(* IEC 61131-3 sources: traffic-lights/PLC_TrafficLights/Class/SafetyManager (part 4) *)

          pHelpSafety^.pThis^.NewInst(pPara, pResult);

          IsDestDomain := TRUE;
          return;
        end_if;

        pHelpSafety := pHelpSafety^.pNext;
      end_while;
    end_if;
  end_if;

END_FUNCTION

FUNCTION SafetyManager::PDOLengthCorrection
  VAR
    pHelpConfig : ^t_CfgListElem;
    pHelpPDO    : ^t_PdoListElem;
    pHelpModule : ^t_ModuleListElem;
    pHelpSearchConfig : ^t_CfgListElem;
    FoundIt : BOOL;
    GotFirst : BOOL;
  END_VAR

  // with FSoE we use connections instead of the PDOs (PDOs are only remembered to check the optional state)
  if b_GotFSoEModules then
    return;
  end_if;

  GotFirst := FALSE;

  // check if there is a PDO with a zero length
  pHelpConfig := pConfigs;
  while pHelpConfig do
    pHelpPDO := pHelpConfig^.pFirstPdoCfg;
    while pHelpPDO do
      // remember the first PDO found as our act (to start from)
      if GotFirst = FALSE then
        GotFirst := TRUE;

        pActualSendCfg := pHelpConfig;
        pActualSendPDO := pHelpPDO;
      end_if;

      // if there is a PDO with no length
      if pHelpPDO^.PdoInfo.PdoLen = 0 then
        FoundIt := FALSE;
        pHelpSearchConfig := pConfigs;
        // search for the source module, because we use the length of it
        while pHelpSearchConfig & (FoundIt = FALSE) do
          pHelpModule := pHelpSearchConfig^.pFirstModuleCfg;
          while pHelpModule & (FoundIt = FALSE) do
            if pHelpModule^.ModuleInfo.PathLen = pHelpPDO^.PdoInfo.SourcePathLen then
              if (To_StdLib.MemCmp(pHelpModule^.ModuleInfo.pPath, pHelpPDO^.PdoInfo.pSourcePath, pHelpModule^.ModuleInfo.PathLen) = 0) then
                pHelpPDO^.PdoInfo.PdoLen := pHelpModule^.ModuleInfo.PdoOutLen;
                FoundIt := TRUE;
              end_if;
            end_if;

            pHelpModule := pHelpModule^.pNext;
          end_while;

          pHelpSearchConfig := pHelpSearchConfig^.pNext;
        end_while;
      end_if;

      pHelpPDO := pHelpPDO^.pNext;
    end_while;

    pHelpConfig := pHelpConfig^.pNext;
  end_while;

END_FUNCTION

FUNCTION SafetyManager::DoublePDOEntry
  VAR_INPUT
    NewPDO 	: t_PdoCfg;
    pNewCfg 	: ^t_CfgListElem;
  END_VAR
  VAR_OUTPUT
    IsDoubleEntry 	: BOOL;
  END_VAR
  VAR
    pHelpCfg : ^t_CfgListElem;
    pHelpPdo : ^t_PdoListElem;
  END_VAR

  IsDoubleEntry := FALSE;

  // if it's our first config, there is no chance for a double PDO => check only if not first config
  if pNewCfg <> pConfigs then
    // otherwise: search all prior configs for the same PDO (source and destination path match)
    pHelpCfg := pConfigs;
    while pHelpCfg <> pNewCfg do
      pHelpPdo := pHelpCfg^.pFirstPdoCfg;
      while pHelpPdo do
        if (pHelpPdo^.PdoInfo.SourcePathLen = NewPDO.SourcePathLen) & (pHelpPdo^.PdoInfo.DestPathLen = NewPDO.DestPathLen) &
           (To_StdLib.MemCmp(pHelpPdo^.PdoInfo.pSourcePath, NewPDO.pSourcePath, NewPDO.SourcePathLen) = 0) &
           (To_StdLib.MemCmp(pHelpPdo^.PdoInfo.pDestPath, NewPDO.pDestPath, NewPDO.DestPathLen) = 0) then
          // we found the same PDO in a prior config
          IsDoubleEntry := TRUE;
          return;
        end_if;

        pHelpPdo := pHelpPdo^.pNext;
      end_while;

      pHelpCfg := pHelpCfg^.pNext;
    end_while;
  end_if;

END_FUNCTION

FUNCTION SafetyManager::StoreInterfaceRoutingList
  VAR_INPUT
    pPara 	: ^CmdStruct;
    pResult 	: ^results;
    IsFSoE 	: BOOL;
  END_VAR
  VAR
    pHelpManaging : ^t_ManagingComponent;
    EntryNo       : USINT;
    i             : UDINT;
    pHelp         : ^t_InterfaceFrameInfo;
    ActOffset     : UDINT;
    pHelpFSoE     : ^t_IFConnectionInfo;
    j             : UDINT;
    GenerateNo    : USINT;
    OldFSoENo     : DINT;
  END_VAR

  if IsFSoE then

    // if we already have different data from this management component => delete the old stuff first
    if IFFSoENo then
      OldFSoENo := IFFSoENo$DINT;

      // remove the existing stuff of this managing component
      for i$DINT := (OldFSoENo-1) to 0 by -1 do
        // check if it's from the same managing component
        if aIFFSoEInfos[i].pManaging^.pThis$DINT = pPara^.aPara[2] then
          // remove it

          // move the following blocks over this one (if it's not the last)
          if i$UDINT < IFFSoENo-1 then
            for j := i to (IFFSoENo-2) do
              aIFFSoEInfos[j] := aIFFSoEInfos[j+1];
            end_for;
          end_if;
          IFFSoENo -= 1;
        end_if;
      end_for;
    end_if;

    EntryNo := ((pPara^.aPara[0] - sizeof(t_IFInfoFSoE.IsResponse)) / sizeof(t_IFConnectionInfo))$USINT;
    if (EntryNo + IFFSoENo <= MAX_MODULES_IN_OTHER_DOMAINS) then
      ActOffset := 0;
      pHelpManaging := pFirstManagingInterfaceComponent;
      while pHelpManaging do
        // if we found the sender of this list in our list of interfaceframe components, remember the safety numbers
        if pHelpManaging^.pThis$DINT = pPara^.aPara[2] then
          if EntryNo then

            // set the help pointer to the first entry of the interface frame info array
            pHelpFSoE := pPara^.aPara[1]$^t_IFConnectionInfo + sizeof(BOOL);
            for i := 0 to (EntryNo-1) do
              pHelpManaging^.ModuleInfo[i].SafetyNbr := pHelpFSoE^.SafetyNbr;

              if pHelpFSoE^.Flags.IsMaster then
                pHelpManaging^.ModuleInfo[i].InfoBits.IsFSoEMaster := TRUE;
                pHelpManaging^.ModuleInfo[i].InfoBits.IsFSoESlave  := FALSE;
              else
                pHelpManaging^.ModuleInfo[i].InfoBits.IsFSoEMaster := FALSE;
                pHelpManaging^.ModuleInfo[i].InfoBits.IsFSoESlave  := TRUE;
              end_if;

              // we save the whole info for PDO/SDO routing
              aIFFSoEInfos[IFFSoENo].FromOtherSide := pHelpFSoE^;
              aIFFSoEInfos[IFFSoENo].FromOtherSide.FollowUps := 0; // only relevant for the transfer to this domain
              aIFFSoEInfos[IFFSoENo].pManaging := pHelpManaging;

              IFFSoENo += 1;

              if pHelpFSoE^.FollowUps then
                GenerateNo := pHelpFSoE^.FollowUps;
                for j := 1 to GenerateNo do
                  // we save the whole info for PDO/SDO routing
                  aIFFSoEInfos[IFFSoENo].FromOtherSide := pHelpFSoE^;
                  aIFFSoEInfos[IFFSoENo].FromOtherSide.FollowUps := 0; // only relevant for the transfer to this domain
                  aIFFSoEInfos[IFFSoENo].pManaging := pHelpManaging;

                  IFFSoENo += 1;
                end_for;
              end_if;

              pHelpFSoE += sizeof(t_IFConnectionInfo);
            end_for;
          end_if;

          pHelpManaging^.ModuleNo := EntryNo;

          pHelpManaging^.InfoBits.GotIFInfo := TRUE;
          return;
        end_if;

        pHelpManaging := pHelpManaging^.pNext;
      end_while;
    else
      LogError("@0473 (SafetyManager::StoreInterfaceRoutingList) Invalid size of configuration (FSoE)");
    end_if;
  else
    EntryNo := ((pPara^.aPara[0] - sizeof(t_IFInfo.IsResponse)) / sizeof(t_InterfaceFrameInfo))$USINT;

    if (EntryNo + InterfaceFrameNo <= MAX_MODULES_IN_OTHER_DOMAINS) then
      ActOffset := 0;
      pHelpManaging := pFirstManagingInterfaceComponent;
      while pHelpManaging do
        // if we found the sender of this list in our list of interfaceframe components, remember the safety numbers
        if pHelpManaging^.pThis$DINT = pPara^.aPara[2] then
          if EntryNo then
            // set the help pointer to the first entry of the interface frame info array
            pHelp := pPara^.aPara[1]$^t_InterfaceFrameInfo + sizeof(BOOL);
            for i := 0 to (EntryNo-1) do
              // we save the module info's with the domain interface module for TDO/SDO routing
              pHelpManaging^.ModuleInfo[i] := pHelp^.ModuleInfo;

              // we also save the whole info for PDO routing
              aInterfaceFrameInfos[InterfaceFrameNo] := pHelp^;

              // only for IFs where the communication partner is the source
              if aInterfaceFrameInfos[InterfaceFrameNo].IFPdoLen then
                aInterfaceFrameInfos[InterfaceFrameNo].OffsetInDomainModule := ActOffset;
                ActOffset += aInterfaceFrameInfos[InterfaceFrameNo].IFPdoLen;
              end_if;

              InterfaceFrameNo += 1;

              pHelp += sizeof(t_InterfaceFrameInfo);
            end_for;
          end_if;

          pHelpManaging^.ModuleNo := EntryNo;

          pHelpManaging^.InfoBits.GotIFInfo := TRUE;
          return;
        end_if;

        pHelpManaging := pHelpManaging^.pNext;
      end_while;
    else
      LogError("@0475 (SafetyManager::StoreInterfaceRoutingList) Invalid size of configuration");
    end_if;
  end_if;

END_FUNCTION

FUNCTION SafetyManager::AllInterfaceCfgsArrived
  VAR_OUTPUT
    AllReady 	: BOOL;
  END_VAR
  VAR
    pHelpManaging : ^t_ManagingComponent;
  END_VAR

  AllReady := TRUE;

  // check if we have the safety numbers for every interface managing module in the system
  pHelpManaging := pFirstManagingInterfaceComponent;
  while pHelpManaging do
    if pHelpManaging^.InfoBits.IsSynchron & (pHelpManaging^.InfoBits.GotIFInfo = FALSE) then
      AllReady := FALSE;
      return;
    end_if;

    pHelpManaging := pHelpManaging^.pNext;
  end_while;

END_FUNCTION

FUNCTION SafetyManager::SendInterfaceConfigs
  VAR_INPUT
    DestinationThis 	: pVirtualBase;(* := NIL *)
    IsResponse 	: BOOL;(* := FALSE *)
    IsFSoE 	: BOOL;
  END_VAR
  VAR
    pHelpCfg                  : ^t_CfgListElem;
    pHelpModule               : ^t_ModuleListElem;
    pHelpPdo                  : ^t_PdoListElem;
    pHelpConnection           : ^t_FSoEConnectionDetails;
    MyPara                    : CmdStruct;
    MyResult                  : results;
    TmpIFInfo                 : t_IFInfo;
    ModuleInfoNo              : USINT;
    i                         : UDINT;
    pActCRC                   : ^HDINT;
    TmpIFConn                 : t_IFInfoFSoESend;
    pLastReferenceConnection  : ^t_IFConnectionInfo;
  END_VAR

  // collect the safety numbers of this system
  ModuleInfoNo := 0;

  if IsFSoE then
    //reset memory => now 0 is an invalid safety number (= unused element of the array)
    _memset(dest:=#TmpIFConn, usByte:=0, cntr:=sizeof(t_IFInfoFSoESend));
    TmpIFConn.IsResponse := IsResponse;

    pLastReferenceConnection  := NIL;

    // if not all configs available, create and send the available data
    if (LocalCPUCfgNo <> LocalCPUNo) then
      // check FSoE Connections in the available configs
      pHelpCfg := pConfigs;
      while pHelpCfg do
        pHelpConnection := pHelpCfg^.pFirstFSoEConnection;
        while pHelpConnection do
          // only interface connections are relevant
          if pHelpConnection^.Flags.IsInterfaceConnection then
            if pLastReferenceConnection & (pHelpConnection^.SlaveAddress = pLastReferenceConnection^.SlaveAddress) &
               (pHelpConnection^.Flags.IsMaster = pLastReferenceConnection^.Flags.IsMaster) then
              pLastReferenceConnection^.FollowUps += 1;
            else
              // add the modules to the info message
              TmpIFConn.aConnectionInfos[ModuleInfoNo].Flags            := pHelpConnection^.Flags;
              TmpIFConn.aConnectionInfos[ModuleInfoNo].SlaveAddress     := pHelpConnection^.SlaveAddress;
              TmpIFConn.aConnectionInfos[ModuleInfoNo].SafetyNbr        := pHelpConnection^.OwnerSafetyNbr;
              TmpIFConn.aConnectionInfos[ModuleInfoNo].MasterReadSize   := pHelpConnection^.MasterReadSize;
              TmpIFConn.aConnectionInfos[ModuleInfoNo].MasterWriteSize  := pHelpConnection^.MasterWriteSize;
              TmpIFConn.aConnectionInfos[ModuleInfoNo].FollowUps        := 0;

              // some data are only available at the master
              if pHelpConnection^.Flags.IsMaster then
                // no follow ups for master connections
                pLastReferenceConnection                                := NIL;

                TmpIFConn.aConnectionInfos[ModuleInfoNo].ConnectionID   := pHelpConnection^.ConnectionID;
              else
                // update this value for the next connections with the same settings to save a lot of memory
                pLastReferenceConnection                                := #TmpIFConn.aConnectionInfos[ModuleInfoNo];

                TmpIFConn.aConnectionInfos[ModuleInfoNo].ConnectionID   := 0;
              end_if;

              if pHelpConnection^.SlavePathCompLen & pHelpConnection^.pSlavePathComp then
                TmpIFConn.aConnectionInfos[ModuleInfoNo].InterfaceCRC := (pHelpConnection^.pSlavePathComp$^HDINT + 1)^;
              else
                TmpIFConn.aConnectionInfos[ModuleInfoNo].InterfaceCRC := 0;
              end_if;

              ModuleInfoNo += 1;
            end_if;
          end_if;

          pHelpConnection := pHelpConnection^.pNext;
        end_while;

        pHelpCfg := pHelpCfg^.pNext;
      end_while;
    else
      // check FSoE Connections in the sorted list
      pHelpConnection := pSortedConnections;
      while pHelpConnection do
        // only interface connections are relevant
        if pHelpConnection^.Flags.IsInterfaceConnection then
          if pLastReferenceConnection & (pHelpConnection^.SlaveAddress = pLastReferenceConnection^.SlaveAddress) &
             (pHelpConnection^.Flags.IsMaster = pLastReferenceConnection^.Flags.IsMaster) then
            pLastReferenceConnection^.FollowUps += 1;
          else
            // add the modules to the info message
            TmpIFConn.aConnectionInfos[ModuleInfoNo].Flags            := pHelpConnection^.Flags;
            TmpIFConn.aConnectionInfos[ModuleInfoNo].SlaveAddress     := pHelpConnection^.SlaveAddress;
            TmpIFConn.aConnectionInfos[ModuleInfoNo].SafetyNbr        := pHelpConnection^.OwnerSafetyNbr;
            TmpIFConn.aConnectionInfos[ModuleInfoNo].MasterReadSize   := pHelpConnection^.MasterReadSize;
            TmpIFConn.aConnectionInfos[ModuleInfoNo].MasterWriteSize  := pHelpConnection^.MasterWriteSize;
            TmpIFConn.aConnectionInfos[ModuleInfoNo].FollowUps        := 0;

            // some data are only available at the master
            if pHelpConnection^.Flags.IsMaster then
              // no follow ups for master connections
              pLastReferenceConnection                                := NIL;

              TmpIFConn.aConnectionInfos[ModuleInfoNo].ConnectionID   := pHelpConnection^.ConnectionID;
            else
              // update this value for the next connections with the same settings to save a lot of memory
              pLastReferenceConnection                                := #TmpIFConn.aConnectionInfos[ModuleInfoNo];

              TmpIFConn.aConnectionInfos[ModuleInfoNo].ConnectionID   := 0;
            end_if;

            if pHelpConnection^.SlavePathCompLen & pHelpConnection^.pSlavePathComp then
              TmpIFConn.aConnectionInfos[ModuleInfoNo].InterfaceCRC := (pHelpConnection^.pSlavePathComp$^HDINT + 1)^;
            else
              TmpIFConn.aConnectionInfos[ModuleInfoNo].InterfaceCRC := 0;
            end_if;

            ModuleInfoNo += 1;
          end_if;
        end_if;

        pHelpConnection := pHelpConnection^.pNextSorted;
      end_while;
    end_if;

    CheckLocalSlaveAddresses();

    if b_AllLocalSlaveAddressesValid then
      MyPara.uiCmd := CMD_SM_IF_MODULE_INFO_FSOE_OK;
    else
      MyPara.uiCmd := CMD_SM_IF_MODULE_INFO_FSOE;
    end_if;

    MyPara.aPara[0] := ModuleInfoNo * sizeof(t_IFConnectionInfo) + sizeof(t_IFInfoFSoE.IsResponse);
    MyPara.aPara[1] := (#TmpIFConn)$DINT;
  else
    // browse through the configs
    TmpIFInfo.IsResponse := IsResponse;

    pHelpCfg := pConfigs;
    while pHelpCfg do
      pHelpPdo := pHelpCfg^.pFirstPdoCfg;
      while pHelpPdo do
        // if it's a interface broadcast
        if pHelpPdo^.PdoInfo.Info.IFBroadCast then
          // search for the source module
          pHelpModule := pHelpCfg^.pFirstModuleCfg;
          while pHelpModule do
            // if it's an interface source and the interface CRC matches the one of our PDO => Bingo! But to be sure we check also the path length and the path itself
            if pHelpModule^.ModuleInfo.Info.IsInterfaceSource & (pHelpModule^.ModuleInfo.InterfaceCRC = pHelpPdo^.PdoInfo.InterfaceCRC) &
              (pHelpModule^.ModuleInfo.PathLen = pHelpPdo^.PdoInfo.SourcePathLen) &
              (To_StdLib.MemCmp(pHelpModule^.ModuleInfo.pPath, pHelpPdo^.PdoInfo.pSourcePath, pHelpPdo^.PdoInfo.SourcePathLen) = 0) then

              TmpIFInfo.aModuleInfos[ModuleInfoNo].InterfaceCRC          := pHelpModule^.ModuleInfo.InterfaceCRC;
              TmpIFInfo.aModuleInfos[ModuleInfoNo].IFPdoLen              := pHelpPdo^.PdoInfo.PdoLen;
              TmpIFInfo.aModuleInfos[ModuleInfoNo].OffsetInDomainModule  := 0; // the correct offset is calculated in the receiver
              TmpIFInfo.aModuleInfos[ModuleInfoNo].ModuleInfo.SafetyNbr  := pHelpModule^.ModuleInfo.SafetyNbr;

              ModuleInfoNo += 1;
            end_if;

            pHelpModule := pHelpModule^.pNext;
          end_while;
        end_if;

        pHelpPdo := pHelpPdo^.pNext;
      end_while;

      // check the modules of the actual config if there are interface frame destinations (needed for unidirectional communication, otherwise the SDO routing would fail)
      pHelpModule := pHelpCfg^.pFirstModuleCfg;
      while pHelpModule do
        // if it's a interface destination
        if pHelpModule^.ModuleInfo.Info.IsInterfaceDest then
          pActCRC := pHelpModule^.ModuleInfo.pDestCRCs;
          for i := 0 to (pHelpModule^.ModuleInfo.DestCRCNo-1) do
            TmpIFInfo.aModuleInfos[ModuleInfoNo].InterfaceCRC          := pActCRC^;
            TmpIFInfo.aModuleInfos[ModuleInfoNo].IFPdoLen              := 0; // we don't know the length here, we're only the receiver
            TmpIFInfo.aModuleInfos[ModuleInfoNo].OffsetInDomainModule  := 0; // the correct offset is calculated in the receiver
            TmpIFInfo.aModuleInfos[ModuleInfoNo].ModuleInfo.SafetyNbr  := pHelpModule^.ModuleInfo.SafetyNbr;
            TmpIFInfo.aModuleInfos[ModuleInfoNo].ModuleInfo.InfoBits$UDINT := 0;

            pActCRC += sizeof(HDINT);
            ModuleInfoNo += 1;
          end_for;
        end_if;

        pHelpModule := pHelpModule^.pNext;
      end_while;

      pHelpCfg := pHelpCfg^.pNext;
    end_while;

    MyPara.uiCmd := CMD_SM_IF_MODULE_INFO;
    MyPara.aPara[0] := ModuleInfoNo * sizeof(t_InterfaceFrameInfo) + sizeof(TmpIFInfo.IsResponse);
    MyPara.aPara[1] := (#TmpIFInfo)$DINT;
  end_if;

  // if we have only 1 destination => sent it to this destination
  if DestinationThis then
    DestinationThis^.NewInst(#MyPara, #MyResult);
  else
    // otherwise send our safety numbers to every interface managing module in the system
    TellAllInterfaceManagingModules(#MyPara, #MyResult);
  end_if;

END_FUNCTION

FUNCTION SafetyManager::GetIFInfoByCRC
  VAR_INPUT
    InterfaceCRC 	: HDINT;
    pMemOffset 	: ^UDINT;
    pLength 	: ^USINT;
  END_VAR
  VAR_OUTPUT
    SafetyNbr 	: HDINT;
  END_VAR
  VAR
    i : UDINT;
  END_VAR

  SafetyNbr := 0;

  if InterfaceFrameNo then
    for i := 0 to (InterfaceFrameNo-1) do
      // if we found the interface CRC and it's a interface frame we receive (the sender adds the length)
      if (aInterfaceFrameInfos[i].InterfaceCRC = InterfaceCRC) & aInterfaceFrameInfos[i].IFPdoLen then
        SafetyNbr := aInterfaceFrameInfos[i].ModuleInfo.SafetyNbr;
        // check if pointers are valid
        if pMemOffset & pLength then
          pMemOffset^ := aInterfaceFrameInfos[i].OffsetInDomainModule;
          pLength^    := aInterfaceFrameInfos[i].IFPdoLen;
        end_if;
        return;
      end_if;
    end_for;

    if SafetyNbr = 0 then
      LogError("@0476 (SafetyManager::GetIFInfoByCRC) Safetynumber of Interface-Frame source couldn't be found in the list");
    end_if;
  end_if;

END_FUNCTION

FUNCTION SafetyManager::SetTimeout

  ud_InitTimeOut := ops.tAbsolute;

END_FUNCTION

FUNCTION SafetyManager::CheckTimeout

  // if the step took too long
  if (OPS.tAbsolute - ud_InitTimeOut) > T_INIT_TIMEOUT then
    // show the possible error in the log/trace and restart the time for timeout
    case InitSSW of
//**********************************************************************************************************************************************************
      _FirstWait4SynchronSubdomains:
        LogError("@0477 (SafetyManager::CheckTimeout) Timeout in Initialisation while waiting first time for subdomains to get synchron!");
//**********************************************************************************************************************************************************
      _Wait4FSoEConnectionsLocal:
        LogError("@0478 (SafetyManager::CheckTimeout) Timeout in Initialisation while waiting for the local FSoE connections to get initialized!");
//**********************************************************************************************************************************************************
      _Wait4SynchronSubdomains:
        LogError("@0479 (SafetyManager::CheckTimeout) Timeout in Initialisation while waiting for subdomains to get synchron!");
//**********************************************************************************************************************************************************
//      _Wait4ConfigFlush:
//        LogError("@ZZZZ Timeout in Initialisation while waiting for the slave domains to send their safety numbers of safety cpus and if they can handle the new time sync method!");
//**********************************************************************************************************************************************************
      _Wait4CPUConfigs:
        LogError("@047A (SafetyManager::CheckTimeout) Timeout in Initialisation while waiting for all available cpu configurations!");
//**********************************************************************************************************************************************************
      _Wait4InterfaceConfigs:
        LogError("@047B (SafetyManager::CheckTimeout) Timeout in Initialisation while waiting for module info needed for interface frame communication!");
//**********************************************************************************************************************************************************
      _Wait4FSoEConnectionsExternal:
        LogError("@047C (SafetyManager::CheckTimeout) Timeout in Initialisation while waiting for the external FSoE connections to get initialized!");
//**********************************************************************************************************************************************************
      _Wait4UnsafeConfigAck:
        LogError("@047D (SafetyManager::CheckTimeout) Timeout in Initialisation while waiting for an unsafe variable configuration acknowledgment!");
//**********************************************************************************************************************************************************
      _Wait4PDOAcks:
        LogError("@047F (SafetyManager::CheckTimeout) Timeout in Initialisation while waiting for a pdo configuration acknowledgment!");
//**********************************************************************************************************************************************************
    end_case;

    // this error gets quitted if initialisation finishes
    ClassState := -11;

    ud_InitTimeOut := ops.tAbsolute;
  end_if;

END_FUNCTION

FUNCTION SafetyManager::AllNonOptionalIFDomainsSynchron
  VAR_OUTPUT
    EverythingSynchron 	: BOOL;
  END_VAR
  VAR
    pHelpManaging : ^t_ManagingComponent;
    pHelpConfig : ^t_CfgListElem;
    pHelpPdo : ^t_PdoListElem;
    TempCfg : t_PdoCfg;
    MyPara 	  : CmdStruct;
    MyResult	: results;
  END_VAR

  EverythingSynchron := TRUE;

  MyPara.uiCmd := CMD_SM_SYNC_CHECK;

  // check for all interface frame PDOs in the configurations if the corresponding domain managing module is synchron
  pHelpConfig := pConfigs;
  while pHelpConfig do
    pHelpPdo := pHelpConfig^.pFirstPdoCfg;
    while pHelpPdo do
      TempCfg := pHelpPdo^.PdoInfo;
      // if it's an interface  PDO, no double entry and not optional => it has to be synchron!
      if (TempCfg.Info.IsInterfacePDO = TRUE) & (TempCfg.Info.DoublePDOEntry = FALSE) & (TempCfg.Info.IsOptional = FALSE) then
        pHelpManaging := pFirstManagingInterfaceComponent;
        while pHelpManaging do
          // we found the corresponding domain managing module
          if (pHelpManaging^.InfoBits.IsOptional = FALSE) &
            ((To_StdLib.MemCmp(pHelpManaging^.pModulePath, TempCfg.pSourcePath, TempCfg.SourcePathLen) = 0) |
             (To_StdLib.MemCmp(pHelpManaging^.pModulePath, TempCfg.pDestPath, TempCfg.DestPathLen) = 0)) then

            // if any of those is not synchron, stop searching
            if pHelpManaging^.pThis^.NewInst(#MyPara, #MyResult) = ERROR then
              EverythingSynchron := FALSE;
              return;
            end_if;

            exit;
          end_if;

          pHelpManaging := pHelpManaging^.pNext;
        end_while;
      end_if;

      pHelpPdo := pHelpPdo^.pNext;
    end_while;

    pHelpConfig := pHelpConfig^.pNext;
  end_while;

END_FUNCTION

FUNCTION VIRTUAL SafetyManager::GetThisViaServerName
  VAR_INPUT
    pObjectDotServer 	: ^CHAR;
  END_VAR
  VAR_OUTPUT
    ThisPtr 	: pVoid;
  END_VAR
  VAR
    ChannelMode : CHMODE;
  END_VAR

  ThisPtr := NIL;

  if pObjectDotServer = NIL then
    return;
  end_if;

  // get thispointer to server via name
  ChannelMode := _LookUpEmbed_C(pObjectDotServer, #ThisPtr, NIL);

  // check if it's a server
  case ChannelMode of
    _CH_CMD,
    _CH_SVR:

  else
    ThisPtr := NIL;
    LogError("@0480 (SafetyManager::GetThisViaServerName) Couldn't get thispointer of server:");
    LogError(e_msg:=pObjectDotServer);
  end_case;

END_FUNCTION

FUNCTION SafetyManager::GetNewMovDO
  VAR_OUTPUT
    Index 	: INT;
  END_VAR
//  VAR
//  	sd_retval : DINT;
//  END_VAR

  Index := -1;

  if CopyCmdsUsed < MAX_PDO_COPY_CMDS then
    // check if there is one available but not used
    if CopyCmdsUsed < CopyCmdsAvailable then
      Index := CopyCmdsUsed;
      CopyCmdsUsed += 1;
    else
      // we have to create a new one

(*
// connection to varan manager required
      // add data object to copy our data
      sd_retval := pVaranManager^.AddMovDO(ud_dol_type:=VARAN_DOL_ISO
                                         , p_ud_handle:=(#aCopyCmds[CopyCmdsAvailable].pHandle)$^UDINT
                                         , p_ud_MovSettings:=( #aCopyCmds[CopyCmdsAvailable].pSettings)$^UDINT
                                         , ud_type := VM_PRIORITY_2
                                         );

      //look for an error
      if ( sd_retval <> 0 ) then
        ClassState := -9;
        LogError("@ZZZZ (SafetyManager::GetNewMovDO) Failed to add a new copy command to the VaranManager!");
        return;
      end_if;
*)
      aCopyCmds[CopyCmdsAvailable].b_Ready4Action := FALSE;

      Index := CopyCmdsAvailable;

      CopyCmdsAvailable += 1;
      CopyCmdsUsed += 1;
    end_if;
  else
    LogError("@0481 (SafetyManager::GetNewMovDO) Maximum of possible PDO copy commands reached!");
  end_if;

END_FUNCTION

FUNCTION SafetyManager::CheckCPUConfigs
  VAR_OUTPUT
    ConfigsOK 	: BOOL;
  END_VAR
  VAR
    pHelpManaging   : ^t_ManagingComponent;
    pSourceManaging : ^t_ManagingComponent;
    pHelpConfig     : ^t_CfgListElem;
    pHelpPdo        : ^t_PdoListElem;
    pLastPdo        : ^t_PdoListElem;
    IsSource        : DINT;
    PDOCount : UDINT;
  END_VAR

  // before we go into the usual check routine, we have to ensure that we have enough virtual PDOs for writing interface frames (config holds a broadcast and we have to look for possible target modules)
  CreateVirtualPDOs();

  // initialize with true (normal case is that everything is ok => now we check for errors)
  ConfigsOK := TRUE;

  PDOCount := 0;

  // check if all non-optional modules are available and all corresponding domain managing module are synchron (if necessary)
  pHelpConfig := pConfigs;
  while pHelpConfig do
    pLastPdo := NIL;
    pHelpPdo := pHelpConfig^.pFirstPdoCfg;
    while pHelpPdo do
      // if it's an interface frame and no broadcast frame
      if pHelpPdo^.PdoInfo.Info.IsInterfacePDO then
        if (pHelpPdo^.PdoInfo.Info.IFBroadCast = FALSE) then

          // check if we have already added the domain interface to the IF List
          IsSource := -1; // -1 = not found, 0 = destination, 1 = source
          pSourceManaging := NIL;
          pHelpManaging := pFirstManagingInterfaceComponent;
          while pHelpManaging do
            // if source or destination of the PDO matches our managing module path => it's an interface frame to/from this domain
            if (To_StdLib.MemCmp(pHelpManaging^.pModulePath, pHelpPdo^.PdoInfo.pSourcePath, pHelpPdo^.PdoInfo.SourcePathLen) = 0) then
              pSourceManaging := pHelpManaging;
              IsSource := 1;
              exit;
            elsif (To_StdLib.MemCmp(pHelpManaging^.pModulePath, pHelpPdo^.PdoInfo.pDestPath, pHelpPdo^.PdoInfo.DestPathLen) = 0) then
              IsSource := 0;
              exit;
            end_if;

            pHelpManaging := pHelpManaging^.pNext;
          end_while;

          // if we got a source managing module and it isn't synchron
          if pSourceManaging then
            // if this pdo is not optional => the source module also isn't
            if pHelpPdo^.PdoInfo.Info.IsOptional = FALSE then
              pSourceManaging^.InfoBits.IsOptional := FALSE;
            end_if;

            if (pSourceManaging^.InfoBits.IsSynchron = FALSE) then
              if pHelpPdo^.PdoInfo.Info.IsOptional then
                // ignore it
  //              LogError("Info: Optional interface frame can't be received, because source domain is not connected or not synchron");

                // remove the PDO from the list (if not the receiver module would wait endless for the PDO and we can't send the set bus ready to quit errors of local PDOs)
                if pLastPdo then
                  // if we had already a PDO before in this configuration we have to skip the removed PDO with the next pointer
                  pLastPdo^.pNext := pHelpPdo^.pNext;

                  To_StdLib.Free(pHelpPdo^.PdoInfo.pSourcePath);
                  To_StdLib.Free(pHelpPdo^.PdoInfo.pDestPath);
                  To_StdLib.Free(pHelpPdo);

                  pHelpPdo := pLastPdo;
                else
                  // if it was the first PDO, we have to correct the first pointer
                  pHelpConfig^.pFirstPdoCfg := pHelpPdo^.pNext;

                  To_StdLib.Free(pHelpPdo^.PdoInfo.pSourcePath);
                  To_StdLib.Free(pHelpPdo^.PdoInfo.pDestPath);
                  To_StdLib.Free(pHelpPdo);

                  pHelpPdo := pHelpConfig^.pFirstPdoCfg;
                end_if;

                if pHelpPdo = NIL then
                  exit;
                end_if;
              else
                // non-optional interface frame domain missing => error
                LogError("@0482 (SafetyManager::CheckCPUConfigs) ERROR! Non-Optional interface frame can't be received, because domain is not connected");
                ConfigsOK := FALSE;
                ClassState := -10;
              end_if;
            end_if;
          end_if;
        end_if;
      end_if;

      PDOCount += 1;

      pLastPdo := pHelpPdo;
      pHelpPdo := pHelpPdo^.pNext;
    end_while;

    pHelpConfig := pHelpConfig^.pNext;
  end_while;

  // if now PDOs found => reset the act ID to show that there are none
  if PDOCount = 0 then
    ActPDO_ID := 0;
  end_if;

END_FUNCTION

FUNCTION SafetyManager::RemoveLocalCPUCfg
  VAR_INPUT
    SafetyNumber 	: HDINT;
  END_VAR
  VAR
    pHelpCfg    : ^t_LocalCfgListElem;
    i : UDINT;
  END_VAR

  if LocalCPUCfgNo then
    pHelpCfg := pFirstLocalCPUCfg;
    for i := 0 to (LocalCPUCfgNo-1) do
      if pHelpCfg^.SafetyNbr = SafetyNumber then
        // found it => deactivate it
        pHelpCfg^.ConfigSize := 0;
        pHelpCfg^.ConfigSent2Master := FALSE;
        exit;
      end_if;

      pHelpCfg := pHelpCfg^.pNext;
    end_for;
  end_if;

END_FUNCTION

FUNCTION SafetyManager::ClearRoutingInformations
  VAR_OUTPUT
    finished 	: BOOL;
  END_VAR
  VAR
    MyPara        : CmdStruct;
    MyResult      : results;
    pHelpManaging : ^t_ManagingComponent;
    i             : UDINT;
    pHelpCfg      : ^t_LocalCfgListElem;
    pPDOElement   : ^t_PDOElement;
    pInputPDO     : ^t_InputPDOs;
    retcode       : DINT;
    pActConnection: ^t_UdpConnection;
    pUdpNo        : ^UDINT;
    paUdpCons     : ^t_aUdpConnections;
  END_VAR

  finished := FALSE;

  if sUdpVars.ProducerConnectionNo then
    pUdpNo    := #sUdpVars.ProducerConnectionNo;
    paUdpCons := sUdpVars.paConnectionsToProducers;
  elsif sUdpVars.ConsumerConnectionNo then
    pUdpNo    := #sUdpVars.ConsumerConnectionNo;
    paUdpCons := sUdpVars.paConnectionsToConsumers;
  else
    // no UDP connections => proceed to last step
    sUdpVars.ClearRoutingInfoSSW := t_ClearRoutingInfoSSW::_FinishEverythingElse;
  end_if;

  case sUdpVars.ClearRoutingInfoSSW of
//**********************************************************************************************************************************************************
    t_ClearRoutingInfoSSW::_PrepareUdpDisconnect:
      // reset all send markers, because we will need them in the next step
      pActConnection := #paUdpCons^[0];
      for i := 0 to (pUdpNo^-1) do
        pActConnection^.WaitForResponse      := FALSE;
        pActConnection^.bSequenceCntReceived := FALSE; //reset flag to allow sequence counter for new udp communication
        pActConnection^.ActReceiveData.usHeaderVersion := 0;
        pActConnection^.ActSendData.usHeaderVersion    := 0;
        pActConnection^.RequestRetries                 := 0;

        pActConnection += sizeof(t_UdpConnection);
      end_for;

      sUdpVars.ClearRoutingInfoSSW := t_ClearRoutingInfoSSW::_SendDisconnect;

//**********************************************************************************************************************************************************
    t_ClearRoutingInfoSSW::_SendDisconnect:

      // if it's the source of the reinit => don't send him the info, just remove from the list
      if (paUdpCons^[pUdpNo^-1].IP = 0) | (paUdpCons^[pUdpNo^-1].IP = sUdpVars.ReInitSenderIP) then
        pUdpNo^ -= 1;
      else
        // disconnect all UDP connections (1 by 1 or we might get a problem with the net load)
        sUdpVars.pTempSendBufferCy^.Header.Command       := t_UdpCommand::UdpCmd_ReInitialize;
        sUdpVars.pTempSendBufferCy^.Header.State         := t_UdpPacketHeaderV2.State.IsFromConsumer OR t_UdpPacketHeaderV2.State.IsFromProducer; // invalid state for normal data

        paUdpCons^[pUdpNo^-1].InfoBits.Disconnecting  := TRUE;
        paUdpCons^[pUdpNo^-1].WaitForResponse         := TRUE;
        paUdpCons^[pUdpNo^-1].TLastRequest            := ops.tAbsolute;

        // only send command and state
        retcode := SendUDPData(sUdpVars.pTempSendBufferCy, sizeof(t_UdpPacketHeaderV2.Command) + sizeof(t_UdpPacketHeaderV2.State), paUdpCons^[pUdpNo^-1].IP);

        if retcode < 0 then
          sUdpVars.LastSendError := retcode;
          sUdpVars.SendErrorCnt += 1;
        end_if;

        sUdpVars.ClearRoutingInfoSSW := t_ClearRoutingInfoSSW::_Wait4DisconnectConfirm;
      end_if;

//**********************************************************************************************************************************************************
    t_ClearRoutingInfoSSW::_Wait4DisconnectConfirm:

      // check for the confirmation
      if paUdpCons^[pUdpNo^-1].InfoBits.Disconnecting = FALSE then

        // reset the IP address of all others with the same IP to not resend if there are multiple connections to this IP
        if sUdpVars.ConsumerConnectionNo then
          pActConnection := #sUdpVars.paConnectionsToConsumers^[0];
          for i := 0 to (sUdpVars.ConsumerConnectionNo-1) do
            // check if it's the same IP
            if (pActConnection^.IP = paUdpCons^[pUdpNo^-1].IP) then
              // reset the IP
              pActConnection^.IP := 0;
            end_if;

            pActConnection += sizeof(t_UdpConnection);
          end_for;
        end_if;

        if sUdpVars.ProducerConnectionNo then
          pActConnection := #sUdpVars.paConnectionsToProducers^[0];
          for i := 0 to (sUdpVars.ProducerConnectionNo-1) do
            // check if it's the same IP
            if (pActConnection^.IP = paUdpCons^[pUdpNo^-1].IP) then
              // reset the IP
              pActConnection^.IP := 0;
            end_if;

            pActConnection += sizeof(t_UdpConnection);
          end_for;
        end_if;

        // this one is out fine => proceed with the next
        pUdpNo^ -= 1;
        sUdpVars.ClearRoutingInfoSSW := t_ClearRoutingInfoSSW::_SendDisconnect;

      // look if we actual wait for a response to send retries and check if we didn't receive data in time
      elsif (paUdpCons^[pUdpNo^-1].WaitForResponse = TRUE) & ((ops.tAbsolute - paUdpCons^[pUdpNo^-1].TLastRequest) > (sUdpVars.CalculatedRequestTimeout * 2)) then

        if paUdpCons^[pUdpNo^-1].RequestRetries >= (UDP_MAX_RETRIES * 2) then

          // we had enough retries, just forget about this one and proceed with the next
          pUdpNo^ -= 1;
          sUdpVars.ClearRoutingInfoSSW := t_ClearRoutingInfoSSW::_SendDisconnect;
        else

          //send retry to actual cpu
          paUdpCons^[pUdpNo^-1].RequestRetries += 1;
          sUdpVars.ClearRoutingInfoSSW := t_ClearRoutingInfoSSW::_SendDisconnect;
        end_if;

      end_if;

      // producer finished but still some consumer connections to go
      if (pUdpNo^ = 0) then
        if sUdpVars.ConsumerConnectionNo then
          // go back to the initialisation and do it for the consumer connections now
          sUdpVars.ClearRoutingInfoSSW := t_ClearRoutingInfoSSW::_PrepareUdpDisconnect;
        else
          // all connections disconnected => finish the rest
          sUdpVars.ClearRoutingInfoSSW := t_ClearRoutingInfoSSW::_FinishEverythingElse;
        end_if;
      end_if;

//**********************************************************************************************************************************************************
    t_ClearRoutingInfoSSW::_FinishEverythingElse:

      // we're flushin our stuff here

      // forget who sent us the reinitialize
      sUdpVars.ReInitSenderIP := 0;

      // set ID to zero for the next mapping assignment
      ActPDO_ID := 0;

      // reset interface frameno
      InterfaceFrameNo := IFFSoENo := 0;

      // reset local interface frameno
      LocalIFNo := 0;

      // clear configurations of safety-cpus
      FreeCfgLists();

      // clear number of copy DOs used
      CopyCmdsUsed := 0;

      // reset flexible constellation informations
      _memset(dest:=#sFlexCon, usByte:=0, cntr:=sizeof(t_FlexCon));

      // reset memory usage for isochronous transfer (the values are set when distributing the PDOs)
      MyPara.aPara[0] := 0;
      pHelpManaging := pFirstManagingInterfaceComponent;
      while pHelpManaging do
        pHelpManaging^.PDOReadMemUsed := 0;
        pHelpManaging^.PDOWriteMemUsed := 0;

        MyPara.uiCmd := CMD_SM_PDO_MEM_USAGE_WR;
        pHelpManaging^.pThis^.NewInst(#MyPara, #MyResult);

        MyPara.uiCmd := CMD_SM_PDO_MEM_USAGE_RD;
        pHelpManaging^.pThis^.NewInst(#MyPara, #MyResult);

        pHelpManaging^.InfoBits.HasBeenFlushed      := FALSE;
        pHelpManaging^.InfoBits.NewTimeSyncPossible := FALSE;
        pHelpManaging^.InfoBits.SubDomainsSynchron  := FALSE;
        pHelpManaging^.InfoBits.GotIFInfo           := FALSE;
        pHelpManaging^.InfoBits.LocalConfigReady    := FALSE;
        pHelpManaging^.InfoBits.IsOptional          := TRUE;  // initialize with true, later in the init process (CheckCPUConfigs) it's checked and corrected if necessary
        // synchron bit is already true at this time (or the timeout has expired)

        pHelpManaging^.DomainNr := 16#FF;

        pHelpManaging^.SubDomainsUsed := 0;
        _memset(dest:=#pHelpManaging^.SubDomainNr, usByte:=16#FF, cntr:=sizeof(pHelpManaging^.SubDomainNr));

        pHelpManaging^.ModuleNo := 0;
        _memset(dest:=#pHelpManaging^.ModuleInfo, usByte:=16#00, cntr:=sizeof(pHelpManaging^.ModuleInfo));

        // delete flexcon information
        _memset(dest:=#pHelpManaging^.FlexCon, usByte:=0, cntr:=sizeof(t_ManagingFlexCon));

        pHelpManaging := pHelpManaging^.pNext;
      end_while;

      // all local cpu configs have to be sent again on reconnect
      if LocalCPUCfgNo then
        pHelpCfg := pFirstLocalCPUCfg;
        for i := 0 to (LocalCPUCfgNo-1) do
          pHelpCfg^.ConfigSent2Master := FALSE;

          pHelpCfg := pHelpCfg^.pNext;
        end_for;
      end_if;

      if PDOElementNo then

        // at first we have to check if there are any safety modules out there with a pointer to the PDO List (if they use a VMC/VBC as source)
        pPDOElement := #aPDOElements[0];
        for i := 0 to (PDOElementNo-1) do
          if (pPDOElement^.ThisDomainsRole = SourceDest_IsDest) & (pPDOElement^.SourceInfo.pPDOMem) & (pPDOElement^.pSafety) then
            // unregister this PDO
            MyPara.uiCmd := CMD_SM_REMOVE_INPUT_PDO;
            MyPara.aPara[0] := pPDOElement^.SourceInfo.pPDOMem$DINT;
            MyPara.aPara[1] := pPDOElement^.SourceInfo.pPDOMemDPRAM$DINT;
            pPDOElement^.pSafety^.pThis^.NewInst(#MyPara, #MyResult);
          end_if;

          // free the memory of the path infos and reset the rest of pdo element info
          if pPDOElement^.SourceInfo.pPath then
            To_StdLib.Free(pPDOElement^.SourceInfo.pPath);
          end_if;
          if pPDOElement^.DestInfo.pPath then
            To_StdLib.Free(pPDOElement^.DestInfo.pPath);
          end_if;

          pPDOElement += sizeof(t_PDOElement);
        end_for;

        _memset(dest:=#aPDOElements, usByte:=0, cntr:=PDOElementNo * sizeof(t_PDOElement));
        PDOElementNo := 0;
      end_if;

      if FSoECopyCmdNo then
        _memset(dest:=#aFSoECopyCmds, usByte:=0, cntr:=FSoECopyCmdNo * sizeof(t_FSoECopyCmd));
        FSoECopyCmdNo := 0;
      end_if;

      if FSoEInputPDONo then
        pInputPDO := #aFSoEInputPDOs[0];
        for i := 0 to (FSoEInputPDONo-1) do
          // unregister this PDO
          MyPara.uiCmd := CMD_SM_REMOVE_INPUT_PDO;
          MyPara.aPara[0] := pInputPDO^.pMem;
          MyPara.aPara[1] := 0;
          pInputPDO^.pSafety^.pThis^.NewInst(#MyPara, #MyResult);

          pInputPDO += sizeof(t_InputPDOs);
        end_for;

        FSoEInputPDONo := 0;
      end_if;

      // reset other udp settings that are not directly connected to the udp connections
      sUdpVars.UdpInit.ProvidesIF            := 0; // no need to install callback twice and FSoE is still available if it was before
      sUdpVars.LowestTransmissionTime_ms  := UDP_DEFAULT_TRANSMISSION_TIME;
      sUdpVars.ConnectionsInitialized     := FALSE;

      // set scheduler to default until a connection is established
      SetUdpSchedulerGrid();

      if sUdpVars.SendCopyCmdNo then
        _memset(dest:=#sUdpVars.aSendCopyCmds, usByte:=0, cntr:=sUdpVars.SendCopyCmdNo * sizeof(t_FSoECopyCmd));
        sUdpVars.SendCopyCmdNo := 0;
      end_if;

      if sUdpVars.ReceiveCopyCmdNo then
        _memset(dest:=#sUdpVars.aReceiveCopyCmds, usByte:=0, cntr:=sUdpVars.ReceiveCopyCmdNo * sizeof(t_FSoECopyCmd));
        sUdpVars.ReceiveCopyCmdNo := 0;
      end_if;

      // reset step
      sUdpVars.ClearRoutingInfoSSW := t_ClearRoutingInfoSSW::_PrepareUdpDisconnect;

      finished := TRUE;

  end_case;

END_FUNCTION

FUNCTION SafetyManager::CheckPDORecycle
  VAR_INPUT
    SourceDest 	: t_SourceDest;
    pNewPDO 	: ^t_PDOElement;
  END_VAR
  VAR_OUTPUT
    pRecyclePDO 	: ^t_PDOElement;
  END_VAR
  VAR
    i : UDINT;
    pHelpInfo : ^t_PDOModuleInfo;
    pSearchInfo : ^t_PDOModuleInfo;
    ppHelpManaging : ^t_pManagingComponent;
    pSearchManaging : ^t_ManagingComponent;
  END_VAR

  // initialize with invalid
  pRecyclePDO := NIL;

  // if we have no pdoelements yet, quit
  if PDOElementNo = 0 then
    return;
  end_if;

  // we search for a PDO with the same source (then it contains the same data)
  pHelpInfo := #aPDOElements[0].SourceInfo;
  pSearchInfo := #pNewPDO^.SourceInfo;

  case SourceDest of
    SourceDest_IsSource:
      ppHelpManaging := #aPDOElements[0].pManagingSource;
      pSearchManaging := pNewPDO^.pManagingSource;
    SourceDest_IsDest:
      ppHelpManaging := #aPDOElements[0].pManagingDest;
      pSearchManaging := pNewPDO^.pManagingDest;
  else
    return;
  end_case;

  // check if we already have the path info of this source/destination
  for i := 0 to (PDOElementNo-1) do
    // if managing node, pathlength and path matches
    if (ppHelpManaging^ = pSearchManaging) & (pHelpInfo^.PathLen = pSearchInfo^.PathLen) & (To_StdLib.MemCmp(pHelpInfo^.pPath, pSearchInfo^.pPath, pHelpInfo^.PathLen) = 0) then
      // we found our PDO to recycle (PDO is already tranferred over this managing node
      pRecyclePDO := #aPDOElements[i];
      return;
    end_if;

    pHelpInfo       += sizeof(t_PDOElement);
    ppHelpManaging  += sizeof(t_PDOElement);
  end_for;

END_FUNCTION

FUNCTION SafetyManager::AddManagingInfo
  VAR_INPUT
    pPara 	: ^CmdStruct;
  END_VAR
  VAR
    pHelpManaging : ^t_ManagingComponent;
  END_VAR

(*
  Parameter description:
  0..pointer to write PDOs in VARAN manager DPRAM
  1..pointer to read PDOs in VARAN manager DPRAM
  2..thispointer of calling class
  3..pointer to write PDOs in internal memory
  4..pointer to read PDOs in internal memory
  5..maximum available space for write PDOs in bytes
  6..maximum available space for read PDOs in bytes
*)

  pHelpManaging := pFirstManagingInterfaceComponent;
  while pHelpManaging do
    if pHelpManaging^.pThis = pPara^.aPara[2]$pVirtualBase then
      exit;
    end_if;

    pHelpManaging := pHelpManaging^.pNext;
  end_while;

  if pHelpManaging then
    pHelpManaging^.pPDOWriteSpaceDPRAM  := pPara^.aPara[0]$^USINT;
    pHelpManaging^.pPDOReadSpaceDPRAM   := pPara^.aPara[1]$^USINT;

    pHelpManaging^.pPDOWriteSpace       := pPara^.aPara[3]$^USINT;
    pHelpManaging^.pPDOReadSpace        := pPara^.aPara[4]$^USINT;

    pHelpManaging^.PDOWriteMemAvailable := pPara^.aPara[5]$UDINT;
    pHelpManaging^.PDOReadMemAvailable  := pPara^.aPara[6]$UDINT;

    pHelpManaging^.ud_HandlePDOWriteSpaceDPRAM  := pPara^.aPara[7]$UDINT;
    pHelpManaging^.ud_HandlePDOReadSpaceDPRAM   := pPara^.aPara[8]$UDINT;

  end_if;

END_FUNCTION

FUNCTION SafetyManager::CheckModuleUsage
  VAR_INPUT
    Length 	: UINT;
    pData 	: ^void;
    IsFSoEConfig 	: BOOL;
  END_VAR
  VAR_OUTPUT
    retcode 	: DINT;
  END_VAR
  VAR
    pDataHelp : ^void;
    i : UDINT;
    TmpPathLen : UINT;
    TempCfgNo : USINT;
    ModuleCfgInfo : t_ModuleCfgInfo;
    PdoCfgInfo : t_PdoCfgInfo;
    TempConnectionNo : UINT;
  END_VAR

(*
    Memory structure:
      4 Byte: SafetyNumber of CPU (is already there from initialisation in CSCP011_IM::InitSafeModule)
      1 Byte: Number of module configurations which are following
      for every module configuration (first is always the CPU itself)
        1 Byte: Info
        4 Byte: Interface Frame Source SafetyNumber (0 if it is no source for interface frames)
        4 Byte: Interface Frame CRC
        1 Byte: Number of destination inferface frame CRCs
        x Byte: Destination interface frame CRCs (number * sizeof(HDINT)
        2 Byte: Length of hardware path
        x Byte (depending on length in the 2 byte before): Hardwarepath
        2 Byte: Length of compressed hardware path
        x Byte (depending on length in the 2 byte before): Compressed Hardwarepath
        1 Byte: PDO out length for this module
      1 Byte: Number of pdo configurations which are following
      for every PDO configuration
        1 Byte: PDO length
        1 Byte: Interface frame info
        4 Byte: Interface CRC
        2 Byte: Length of source hardware path
        x Byte (depending on length in the 2 byte before): Hardwarepath of source
        2 Byte: Length of destination hardware path
        x Byte (depending on length in the 2 byte before): Hardwarepath of destination
      1 Byte: Number of slave configurations which are following
      for every slave configuration
        1 Byte: Info
        4 Byte: InterfaceCRC
        2 Byte: Length of hardware path
        x Byte (depending on length in the 2 byte before): Hardwarepath
        2 Byte: Length of compressed hardware path
        x Byte (depending on length in the 2 byte before): Compressed Hardwarepath

      if IsFSoEConfig = TRUE
      2 Byte: Number of connection infos which are following
      for every FSoE connection info
        2 Byte: ConnectionID
        1 Byte: ConnectionState
        1 Byte: Flags
        4 Byte: Master safety number

only if feature available:
        2 Byte: Transmission time in ms

        2 Byte: Offset where to read from master
        2 Byte: Size of data to read from master (and write to slave)
        2 Byte: Offset where to write to master
        2 Byte: Size of data to write to master (and read from slave)
        2 Byte: SlaveAddress
        2 Byte: Length of slave hardware path
        x Byte (depending on length in the 2 byte before): Slave hardware path
        2 Byte: Length of compressed slave hardware path
        x Byte (depending on length in the 2 byte before): Compressed slave hardware path
        2 Byte: Offset where to read from slave
        2 Byte: Offset where to write to slave
*)

  // check if the configuration is valid (pData <> NIL) & (Length must be at least 4 byte for SafetyNbr + 1 byte module cfg number + 1 byte pdo cfg number + 1 byte slave cfc number)
  if pData & (Length >= 7)  then

    retcode := 0;

    pDataHelp := pData;

    // skip safety number of the safety cpu
    pDataHelp += sizeof(HDINT);

    // number of module configurations which follow now
    TempCfgNo := pDataHelp^$USINT;

    // skip number of module configurations
    pDataHelp += sizeof(USINT);

    // module configurations
    if TempCfgNo then
      for i := 0 to (TempCfgNo-1) do
        // info
        ModuleCfgInfo := pDataHelp^$t_ModuleCfgInfo;

        // skip info
        pDataHelp += sizeof(BSINT);

        // skip safety number of interface frame source
        pDataHelp += sizeof(HDINT);

        // skip interface CRC of interface frame
        pDataHelp += sizeof(HDINT);

        // interface frame destination CRCs
        if ModuleCfgInfo.IsInterfaceDest then
          // number of CRCs
          TmpPathLen := pDataHelp^$USINT;

          // skip number of CRCs
          pDataHelp += sizeof(USINT);

          // skip interface destination CRCs
          pDataHelp += TmpPathLen * sizeof(HDINT);
        end_if;

        // length of hardware path
        TmpPathLen := pDataHelp^$UINT;

        // skip length of hardware path
        pDataHelp += sizeof(UINT);

        SetModuleUsed(PathLen:=TmpPathLen, pPath:=pDataHelp$^USINT, IgnoreOptional:=FALSE, IsOptional:=ModuleCfgInfo.IsOptional, IsInterfaceDomain := FALSE);

        // skip hardware path
        pDataHelp += TmpPathLen;

        // length of compressed hardware path
        TmpPathLen := pDataHelp^$UINT; // save some time with this local variable

        // skip length of compressed hardware path
        pDataHelp += sizeof(UINT);

        // skip compressed hardware path
        pDataHelp += TmpPathLen;

        // skip pdo out length of this module
        pDataHelp += sizeof(USINT);
      end_for;
    end_if;

    // number of Pdo configurations which follow now
    TempCfgNo := pDataHelp^$USINT;

    // skip number of pdo configurations
    pDataHelp += sizeof(USINT);

    // Pdo configurations
    if TempCfgNo then
      for i := 0 to (TempCfgNo-1) do
        // skip pdo length
        pDataHelp += sizeof(USINT);

        // is it an interface pdo?
        PdoCfgInfo := pDataHelp^$t_PdoCfgInfo;

        // skip info
        pDataHelp += sizeof(BSINT);

        // skip interface CRC
        pDataHelp += sizeof(HDINT);

        // length of source hardware path
        TmpPathLen := pDataHelp^$UINT;

        // skip length of source hardware path
        pDataHelp += sizeof(UINT);

        SetModuleUsed(PathLen:=TmpPathLen, pPath:=pDataHelp$^USINT, IgnoreOptional:=FALSE, IsOptional:=PdoCfgInfo.IsOptional, IsInterfaceDomain := PdoCfgInfo.IsInterfacePDO);

        // skip source hardware path
        pDataHelp += TmpPathLen;

        // length of destination hardware path
        TmpPathLen := pDataHelp^$UINT;

        // skip length of destination hardware path
        pDataHelp += sizeof(UINT);

        // a destination module doesn't influence the optional property=> ignore the optional setting
        SetModuleUsed(PathLen:=TmpPathLen, pPath:=pDataHelp$^USINT, IgnoreOptional:=TRUE, IsOptional:=FALSE, IsInterfaceDomain := PdoCfgInfo.IsInterfacePDO);

        // skip destination hardware path
        pDataHelp += TmpPathLen;
      end_for;
    end_if;

    // number of slave configurations which follow now
    TempCfgNo := pDataHelp^$USINT;

    // skip number of slave configurations
    pDataHelp += sizeof(USINT);

    // slave configurations
    if TempCfgNo then
      for i := 0 to (TempCfgNo-1) do
        // skip info
        pDataHelp += sizeof(BSINT);

        // skip InterfaceCRC
        pDataHelp += sizeof(HDINT);

        // length of hardwarepath
        TmpPathLen := pDataHelp^$UINT; // save some time with this local variable

        // skip length of hardwarepath
        pDataHelp += sizeof(UINT);

        // skip hardwarepath
        pDataHelp += TmpPathLen;

        // length of compressed hardwarepath
        TmpPathLen := pDataHelp^$UINT; // save some time with this local variable

        // skip length of compressed hardwarepath
        pDataHelp += sizeof(UINT);

        // skip compressed hardwarepath
        pDataHelp += TmpPathLen;
      end_for;
    end_if;

    // check if it's a FSoE Config
    if IsFSoEConfig then
      // number of connection details which follow now
      TempConnectionNo := pDataHelp^$UINT;
      pDataHelp += sizeof(UINT);

      // if we got connections
      if TempConnectionNo then
        for i := 0 to (TempConnectionNo-1) do
          // connection ID
          pDataHelp += sizeof(UINT);

          // connection state
          pDataHelp += sizeof(USINT);

          // flags
          // Actually, type is 4 bytes in size but for compatibility reasons it is still used as 1 byte. As a result, bits 9-32 are currently not used.
          pDataHelp += sizeof(t_FSoEFlags);

          // master safety number
          pDataHelp += sizeof(HDINT);

          if bdFeatureEnable.TransmissionTimeInConfig then
            // transmission time in ms
            pDataHelp += sizeof(UINT);
          end_if;

          // offset where to read from master
          pDataHelp += sizeof(UINT);

          // size of data to read from master (and write to slave)
          pDataHelp += sizeof(UINT);

          // offset where to write to master
          pDataHelp += sizeof(UINT);

          // size of data to write to master (and read from slave)
          pDataHelp += sizeof(UINT);

          // slave address
          pDataHelp += sizeof(UINT);

          // length of uncompressed slave hardwarepath
          TmpPathLen := pDataHelp^$UINT; // save some time with this local variable
          pDataHelp += sizeof(UINT);

          // uncompressed slave hardwarepath
          pDataHelp += TmpPathLen;

          // length of compressed slave hardwarepath
          TmpPathLen := pDataHelp^$UINT; // save some time with this local variable
          pDataHelp += sizeof(UINT);

          // compressed slave hardwarepath
          pDataHelp += TmpPathLen;

          // offset where to read from master
          pDataHelp += sizeof(UINT);

          // offset where to write to master
          pDataHelp += sizeof(UINT);
        end_for;
      end_if;
    end_if;

    // check if the given size matches the memory structure
    if (pDataHelp$UDINT - pData$UDINT) <> Length then
      LogError("@459 (SafetyManager::CheckModuleUsage) Invalid configuration data given (length doesn't match memory structure)");
      retcode := -3;
      return;
    end_if;
  else
    // invalid configuration
    LogError("@045A (SafetyManager::CheckModuleUsage) Found invalid safety cpu configuration: Pointer or size wrong");
    retcode := -1;
  end_if;

END_FUNCTION

FUNCTION SafetyManager::SetModuleUsed
  VAR_INPUT
    PathLen 	: UINT;
    pPath 	: ^USINT;
    IgnoreOptional 	: BOOL;
    IsOptional 	: BOOL;
    IsInterfaceDomain 	: BOOL;
  END_VAR
  VAR
    pHelpManaging : ^t_ManagingComponent;
    pHelpSafety   : ^t_SafetyComponent;
    i             : UDINT;
    pActConnection: ^t_UdpConnection;
  END_VAR

  // search for the hardware path

  // only possible for UDP connections
  if sUdpVars.ProducerConnectionNo & (pPath^ = INTERFACE_IP_MODE) & (PathLen = UDP_COMP_PATH_LENGTH) then
    pActConnection := #sUdpVars.paConnectionsToProducers^[0];
    for i := 0 to (sUdpVars.ProducerConnectionNo-1) do
      if (pActConnection^.IFCRC = (pPath$^HDINT + 1)^) & (pActConnection^.IP = (pPath$^HDINT + 5)^) then
        // update optional info
        pActConnection^.InfoBits.IsOptional     := IsOptional;
        pActConnection^.InfoBits.OptionalValid  := TRUE;

        return;
      end_if;

      pActConnection += sizeof(t_UdpConnection);
    end_for;

  else

    // start with the safety components
    pHelpSafety := pFirstSafetyComponent;
    while pHelpSafety & pHelpSafety^.pPath do
      // we have 1 byte path length on the safety component but we got a 2 byte path length from the configuration
      // furthermore the pPath string could be over more domains and we have only our local path => check if length is bigger and if there is a domain escape right before the domain number
      if ((pPath^ = pHelpSafety^.pPath^) | ((pPath^ > pHelpSafety^.pPath^) & ((pPath + 1 + pPath^ - pHelpSafety^.pPath^)^ = HWT_ESCAPE_DOMAIN))) &
         (To_StdLib.MemCmp(pHelpSafety^.pPath + 1, pPath + 2 + pPath^ - pHelpSafety^.pPath^, pHelpSafety^.pPath^) = 0) then
        // only set IsOptional to false (has been initialized with true)
        if (IsOptional = FALSE) & (IgnoreOptional = FALSE) then
          pHelpSafety^.InfoBits.IsOptional := FALSE;
        end_if;
        return;
      end_if;

      pHelpSafety := pHelpSafety^.pNext;
    end_while;

    // if not found, continue with the managing interface components
    pHelpManaging := pFirstManagingInterfaceComponent;
    while pHelpManaging do
      if (To_StdLib.MemCmp(pHelpManaging^.pModulePath, pPath, PathLen) = 0) then
        // only set IsOptional to false (has been initialized with true)
        if (IsOptional = FALSE) & (IgnoreOptional = FALSE) then
          pHelpManaging^.InfoBits.IsOptional := FALSE;
        end_if;
        return;
      end_if;

      pHelpManaging := pHelpManaging^.pNext;
    end_while;

  end_if;

END_FUNCTION

FUNCTION SafetyManager::CreateTimeSyncList
  VAR
    pHelp : ^t_TimeSyncElement;
    pHelpSafety   : ^t_SafetyComponent;
    pHelpManaging : ^t_ManagingComponent;
  END_VAR

  // first we stop time syncing (if active) to prevent crashing due tue a running time synchronisation
  pActTimeSyncElement := NIL;

  // if there is an old list, free it first
  if pFirstTimeSyncElement then
    // open the ring (set the next pointer of the last element to NIL)
    pFirstTimeSyncElement^.pPrev^.pNext := NIL;

    // remove the elements
    while pFirstTimeSyncElement do
      pHelp := pFirstTimeSyncElement;
      pFirstTimeSyncElement := pFirstTimeSyncElement^.pNext;

      To_StdLib.Free(mptr:=pHelp);
    end_while;
  end_if;

  pHelpSafety := pFirstSafetyComponent;
  while pHelpSafety do
    // if it's a module with not only inputs (then there's nothing to synchronize with) => trigger it for time synchronisation
    if (pHelpSafety^.InfoBits.OnlyInputs = FALSE) & (IsFSoEModule(pHelpSafety^.ModuleType) = FALSE) then
      AddTimeSyncElement(pManaging:=NIL, pSafety:=pHelpSafety, IsInterfaceDomain := FALSE);
    end_if;

    pHelpSafety := pHelpSafety^.pNext;
  end_while;

  // interface domains will not get our token, they got their own
  pHelpManaging := pFirstManagingInterfaceComponent;
  while pHelpManaging do
    AddTimeSyncElement(pManaging:=pHelpManaging, pSafety:=NIL, IsInterfaceDomain := TRUE);

    pHelpManaging := pHelpManaging^.pNext;
  end_while;

END_FUNCTION

FUNCTION SafetyManager::AddTimeSyncElement
  VAR_INPUT
    pManaging 	: ^t_ManagingComponent;
    pSafety 	: ^t_SafetyComponent;
    IsInterfaceDomain 	: BOOL;
  END_VAR
  VAR
    pLast : ^t_TimeSyncElement;
    pHelp : ^t_TimeSyncElement;
  END_VAR

  // first we have to allocate some memory for the new element
  if pFirstTimeSyncElement = NIL then
    pFirstTimeSyncElement$pVoid := To_StdLib.Malloc(size:=sizeof(t_TimeSyncElement));
    pLast := pHelp := pFirstTimeSyncElement;
  else
    // check if we got this already
    pHelp := pFirstTimeSyncElement;
    repeat
      if pSafety & (pHelp^.pSafety = pSafety) then
        // already in list => leave
        return;
      end_if;

      if pManaging & (pHelp^.pManaging = pManaging) then
        // already in list => leave
        return;
      end_if;

      pHelp := pHelp^.pNext;
    until (pHelp = pFirstTimeSyncElement) end_repeat;

    pHelp$pVoid := To_StdLib.Malloc(size:=sizeof(t_TimeSyncElement));
    pLast := pFirstTimeSyncElement^.pPrev;
  end_if;

  if pHelp then
    // close the double linked ring with the new elements
    pFirstTimeSyncElement^.pPrev := pHelp;
    pHelp^.pNext := pFirstTimeSyncElement;

    pHelp^.pPrev := pLast;
    pLast^.pNext := pHelp;

    pHelp^.InfoBits := 0;
    pHelp^.InfoBits.IsInterfaceDomain := IsInterfaceDomain;

    pHelp^.pManaging := pManaging;
    pHelp^.pSafety   := pSafety;

    // managing modules
    if (pManaging <> NIL) then
      pHelp^.InfoBits.IsManagingModule := TRUE;
      pHelp^.pThis := pManaging^.pThis;

      // if it's the master connection
      if pManaging^.InfoBits.IsConnectionToMaster then
        // remember it
        pHelp^.InfoBits.IsConnectionToMaster := TRUE;

        // and make it the end of the list
        pFirstTimeSyncElement := pHelp^.pNext;

        // remember that we got a master connection
        pMasterTimeSyncElement := pHelp;

      elsif pMasterTimeSyncElement then
        // if we're not master and there is already a master time sync element in the list, we have to make it the last element
        pFirstTimeSyncElement := pMasterTimeSyncElement^.pNext;
      end_if;
    else
      // safety modules
      pHelp^.InfoBits.IsManagingModule := FALSE;
      pHelp^.pThis := pSafety^.pThis;

    // insert new safety modules at the beginning (managing modules at the end)
      pFirstTimeSyncElement := pHelp;
    end_if;

  else
    ClassState := -1;
    LogError("@0485 (SafetyManager::AddTimeSyncElement) Failed to allocate memory for a new Element");
  end_if;

END_FUNCTION

FUNCTION SafetyManager::CreateVirtualPDOs
  VAR
    pHelpManaging   : ^t_ManagingComponent;
    pHelpConfig     : ^t_CfgListElem;
    pHelpPdo        : ^t_PdoListElem;
    TempPDO         : t_PdoCfg;
    pSearchConfig   : ^t_CfgListElem;
    pSearchPdo      : ^t_PdoListElem;
    b_UsedAsDest    : BOOL;
  END_VAR

  pHelpConfig := pConfigs;
  while pHelpConfig do
    pHelpPdo := pHelpConfig^.pFirstPdoCfg;
    while pHelpPdo do
      // check if it's a broadcast
      if (pHelpPdo^.PdoInfo.Info.IFBroadCast) & (pHelpPdo^.PdoInfo.Info.VirtualPDOsCreated = FALSE) then
        // found one => create virtual PDOs from it (add them to the same configuration)

        // prepare new virtual PDO
        TempPDO := pHelpPdo^.PdoInfo;

        TempPDO.Info.IFBroadCast := FALSE;
        TempPDO.Info.VirtualPDO := TRUE;

        // add a new PDO for every interface managing module
        pHelpManaging := pFirstManagingInterfaceComponent;
        while pHelpManaging do
          // change destination path to the actual module
          TempPDO.DestPathLen := pHelpManaging^.pModulePath^ + 2;
          TempPDO.pDestPath := pHelpManaging^.pModulePath;

          if AddVirtualPDOToCfg(pCfg:=pHelpConfig, pNewPDO:=#TempPDO) then
            LogError("@0486 (SafetyManager::CreateVirtualPDOs) Failed to allocate memory for a new virtual PDO");
          end_if;

          pHelpManaging := pHelpManaging^.pNext;
        end_while;

        // search in all configs (if there are other) for a pdo with this interface CRC as source
        pSearchConfig := pConfigs;
        while pSearchConfig do
          pSearchPdo := pSearchConfig^.pFirstPdoCfg;
          while pSearchPdo do
            // we must not manipulate our help pdo
            if pSearchPdo <> pHelpPdo then
              b_UsedAsDest := FALSE;

              // check if the path is already used as destination
              if (pSearchPdo^.PdoInfo.DestPathLen = pHelpPdo^.PdoInfo.SourcePathLen) &
                 (To_StdLib.MemCmp(pSearchPdo^.PdoInfo.pDestPath, pHelpPdo^.PdoInfo.pSourcePath, pHelpPdo^.PdoInfo.SourcePathLen) = 0) then
                b_UsedAsDest := TRUE;
              end_if;

              // check if the interface CRC appears in any PDO (only if the path isn't already used as destination path)
              if (pSearchPdo^.PdoInfo.InterfaceCRC = pHelpPdo^.PdoInfo.InterfaceCRC) & (b_UsedAsDest = FALSE) then
                // now take the source path of the broadcast PDO and use it as source path for this PDO
                To_StdLib.Free(mptr:=pSearchPdo^.PdoInfo.pSourcePath);

                pSearchPdo^.PdoInfo.pSourcePath$pVoid := To_StdLib.Malloc(size:=pHelpPdo^.PdoInfo.SourcePathLen);

                // save source hardwarepath
                if pSearchPdo^.PdoInfo.pSourcePath then
                  _memcpy(ptr1:=pSearchPdo^.PdoInfo.pSourcePath, ptr2:=pHelpPdo^.PdoInfo.pSourcePath, cntr:=pHelpPdo^.PdoInfo.SourcePathLen);
                  pSearchPdo^.PdoInfo.SourcePathLen := pHelpPdo^.PdoInfo.SourcePathLen;

                  // source and destination of this PDO are both local safe cpu modules which communicate with each other via interface frames => store them in extra list for routing SDOs and TDOs
                  AddToLocalIFs(#pSearchPdo^.PdoInfo);
                else
                  LogError("@0487 (SafetyManager::CreateVirtualPDOs) Failed to allocate memory for a source path");
                  pSearchPdo^.PdoInfo.SourcePathLen := 0;
                  ClassState := -1;
                end_if;
              end_if;
            end_if;

            pSearchPdo := pSearchPdo^.pNext;
          end_while;

          pSearchConfig := pSearchConfig^.pNext;
        end_while;
        pHelpPdo^.PdoInfo.Info.VirtualPDOsCreated := TRUE;
      end_if;

      pHelpPdo := pHelpPdo^.pNext;
    end_while;

    pHelpConfig := pHelpConfig^.pNext;
  end_while;

END_FUNCTION

FUNCTION SafetyManager::AddVirtualPDOToCfg
  VAR_INPUT
    pCfg 	: ^t_CfgListElem;
    pNewPDO 	: ^t_PdoCfg;
  END_VAR
  VAR_OUTPUT
    retcode 	: DINT;
  END_VAR
  VAR
    pHelpPdo        : ^t_PdoListElem;
    TempLen         : UINT;
  END_VAR

  retcode := 0;

  if pCfg^.pFirstPdoCfg = NIL then
    // first PDO in this cfg (should not be possible, because the template for this PDO is also in the same config)
    pCfg^.pFirstPdoCfg$pVoid := To_StdLib.Malloc(size:=sizeof(t_PdoListElem));
    pHelpPdo := pCfg^.pFirstPdoCfg;
  else
    // search a place for the new PDO
    pHelpPdo := pCfg^.pFirstPdoCfg;
    while pHelpPdo^.pNext do

      pHelpPdo := pHelpPdo^.pNext;
    end_while;

    pHelpPdo^.pNext$pvoid := To_StdLib.Malloc(size:=sizeof(t_PdoListElem));
    pHelpPdo := pHelpPdo^.pNext;
  end_if;

  if pHelpPdo then
    // init the values
    pHelpPdo^.PdoInfo.PdoLen        := pNewPDO^.PdoLen;
    pHelpPdo^.PdoInfo.Info          := pNewPDO^.Info;
    pHelpPdo^.PdoInfo.InterfaceCRC  := pNewPDO^.InterfaceCRC;

    // length of source hardwarepath
    TempLen := pNewPDO^.SourcePathLen; // save some time with this local variable
    pHelpPdo^.PdoInfo.SourcePathLen := TempLen;

    // allocate memory for the source module path
    pHelpPdo^.PdoInfo.pSourcePath$pVoid := To_StdLib.Malloc(size:=TempLen);
    if pHelpPdo^.PdoInfo.pSourcePath = NIL then
      ClassState := -1;
      retcode := -2;
      return;
    end_if;

    // save source hardwarepath
    _memcpy(ptr1:=pHelpPdo^.PdoInfo.pSourcePath, ptr2:=pNewPDO^.pSourcePath, cntr:=TempLen);

    // length of destination hardwarepath
    TempLen := pNewPDO^.DestPathLen; // save some time with this local variable
    pHelpPdo^.PdoInfo.DestPathLen := TempLen;

    // allocate memory for the destination module path
    pHelpPdo^.PdoInfo.pDestPath$pVoid := To_StdLib.Malloc(size:=TempLen);
    if pHelpPdo^.PdoInfo.pDestPath = NIL then
      ClassState := -1;
      retcode := -2;
      return;
    end_if;

    // save destination hardwarepath
    _memcpy(ptr1:=pHelpPdo^.PdoInfo.pDestPath, ptr2:=pNewPDO^.pDestPath, cntr:=TempLen);

    // now we give it an ID and increase the number for the next pdo
    pHelpPdo^.PdoInfo.PDO_ID := ActPDO_ID;
    ActPDO_ID += 1;

    pHelpPdo^.pNext                  := NIL;
  else
    ClassState := -1;
    retcode := -2;
    return;
  end_if;

END_FUNCTION

FUNCTION SafetyManager::AddToLocalIFs
  VAR_INPUT
    pHelpPDO 	: ^t_PdoCfg;
  END_VAR
  VAR
    AddSource : BOOL;
    i : USINT;
    pHelpSafety : ^t_SafetyComponent;
  END_VAR

  // check if there is still room for new modules
  if LocalIFNo < MAX_INTERNAL_IF_MODULES then

    AddSource := TRUE;

    // if there is a list, check if any of our modules are already in the list
    if LocalIFNo then
      for i := 0 to (LocalIFNo-1) do
        // check if crc matches
        if (aLocalIFs[i].InterfaceCRC = pHelpPDO^.InterfaceCRC) then
          AddSource := FALSE;
          exit;
        end_if;
      end_for;
    end_if;

    // now we know how many we have to add to the list. if there are modules to add and there is enough space for all of them => do it
    if AddSource then
      // search it in the local modules
      pHelpSafety := pFirstSafetyComponent;
      while pHelpSafety do
        // if the path matches, add the module to the list

        // source module
        if (pHelpSafety^.PathLen = (pHelpPDO^.SourcePathLen - 1)) &
        // we compare the last x byte (where x is the length of the local path including the domain) because we got different length info sizes (1 byte vs. 2 byte)
           (To_StdLib.MemCmp(pHelpSafety^.pPath + 1, pHelpPDO^.pSourcePath + 2 + pHelpPDO^.pSourcePath^ - pHelpSafety^.pPath^, pHelpSafety^.pPath^) = 0) then
          aLocalIFs[LocalIFNo].InterfaceCRC  := pHelpPDO^.InterfaceCRC;
          aLocalIFs[LocalIFNo].pSafetyModule := pHelpSafety;
          LocalIFNo += 1;
          exit;
        end_if;

        pHelpSafety := pHelpSafety^.pNext;
      end_while;
    end_if;
  end_if;

END_FUNCTION

FUNCTION SafetyManager::IFInfoNotArrivedYet
  VAR_INPUT
    pThis 	: pVirtualBase;
  END_VAR
  VAR_OUTPUT
    InfoNotAvailable 	: BOOL;
  END_VAR
  VAR
    pHelpManaging : ^t_ManagingComponent;
  END_VAR

  InfoNotAvailable := FALSE;

  pHelpManaging := pFirstManagingInterfaceComponent;
  while pHelpManaging do
    if pHelpManaging^.pThis = pThis then
      if pHelpManaging^.InfoBits.GotIFInfo = FALSE then
        InfoNotAvailable := TRUE;
      end_if;
      return;
    end_if;

    pHelpManaging := pHelpManaging^.pNext;
  end_while;

END_FUNCTION

#pragma warning(disable:74)
#pragma warning(disable:73)
FUNCTION SafetyManager::StartTimeMeasurement
  VAR_INPUT
    usMode (EAX) 	: DINT;
  END_VAR
#ifdef VM_CLASS_TIME_MEASUREMENT
  VAR
    tmpTime : ^t_TimeMeasurementVaran;
  END_VAR

  case usMode of

    //-----------------------------------------------------------

    VARANTIME_RT:
      tmpTime := #s_TimeRt;

    //-----------------------------------------------------------

    VARANTIME_RTPOSTSCAN:
      tmpTime := #s_TimeRtPostScan;

    //-----------------------------------------------------------

    VARANTIME_CY:
      tmpTime := #s_TimeCy;

    //-----------------------------------------------------------

  end_case;

  if ( tmpTime^.us_Activate ) then
//    Save_Flg();
//    CLI();
    tmpTime^.ud_Timemark := OS_READMICROSEC();
  end_if;

#endif

END_FUNCTION

FUNCTION SafetyManager::StopTimeMeasurement
  VAR_INPUT
    usMode (EAX) 	: DINT;
  END_VAR
#ifdef VM_CLASS_TIME_MEASUREMENT
  VAR
    tmpTime : ^t_TimeMeasurementVaran;
  END_VAR

  case usMode of

    //-----------------------------------------------------------

    VARANTIME_RT:
      tmpTime := #s_TimeRt;

    //-----------------------------------------------------------

    VARANTIME_RTPOSTSCAN:
      tmpTime := #s_TimeRtPostScan;

    //-----------------------------------------------------------

    VARANTIME_CY:
      tmpTime := #s_TimeCy;

    //-----------------------------------------------------------

  end_case;

  if ( tmpTime^.us_Activate ) then

    //get actual time
    tmpTime^.ud_ActualTime := OS_READMICROSEC();
    tmpTime^.ud_ActualTime -= tmpTime^.ud_Timemark;

    //look for maximum time
    if ( tmpTime^.ud_ActualTime > tmpTime^.ud_MaximalTime ) then
      tmpTime^.ud_MaximalTime := tmpTime^.ud_ActualTime;
    end_if;

    //look for minimum time
    if ( tmpTime^.ud_ActualTime < tmpTime^.ud_MinimalTime ) then
      tmpTime^.ud_MinimalTime := tmpTime^.ud_ActualTime;
    end_if;

    //look for average time (100000 cycles)
    if ( tmpTime^.ud_AverageCounter = 100000 ) then

      tmpTime^.ud_AverageTime 	:= tmpTime^.ud_AverageSum / tmpTime^.ud_AverageCounter;
      tmpTime^.ud_AverageSum 	:= 0;
      tmpTime^.ud_AverageCounter := 0;

    else
      tmpTime^.ud_AverageSum += ( tmpTime^.ud_ActualTime / 100 );
      tmpTime^.ud_AverageCounter += 1;
    end_if;

//		STI();
//    Restore_Flg();
  end_if;

#endif

END_FUNCTION // Varan_Base::StopTimeMeasurement
#pragma warning(default:74)
#pragma warning(default:73)

FUNCTION SafetyManager::AnyIFDomainSynchron
  VAR_OUTPUT
    AnythingSynchron 	: BOOL;
  END_VAR
  VAR
    pHelpManaging   : ^t_ManagingComponent;
  END_VAR

  AnythingSynchron := FALSE;

  pHelpManaging := pFirstManagingInterfaceComponent;
  while pHelpManaging do
    if pHelpManaging^.InfoBits.IsSynchron then
      AnythingSynchron := TRUE;
      return;
    end_if;

    pHelpManaging := pHelpManaging^.pNext;
  end_while;

END_FUNCTION

FUNCTION SafetyManager::LocalIFsAvailable
  VAR_OUTPUT
    retcode 	: BOOL;
  END_VAR
  VAR
    pHelpCfg : ^t_CfgListElem;
    pHelpPdo : ^t_PdoListElem;
    pHelpModule : ^t_ModuleListElem;
  END_VAR

  retcode := FALSE;

  // add all local configs to our structure
  SendLocalCfgsToMaster();

  // check the local configs for interface frames
  pHelpCfg := pConfigs;
  while pHelpCfg do
    pHelpPdo := pHelpCfg^.pFirstPdoCfg;
    while pHelpPdo do
      if pHelpPdo^.PdoInfo.Info.IsInterfacePDO | pHelpPdo^.PdoInfo.Info.IFBroadCast then
        retcode := TRUE;
        return;
      end_if;

      pHelpPdo := pHelpPdo^.pNext;
    end_while;

    pHelpModule := pHelpCfg^.pFirstModuleCfg;
    while pHelpModule do
      if pHelpModule^.ModuleInfo.Info.IsInterfaceSource | pHelpModule^.ModuleInfo.Info.IsInterfaceDest then
        retcode := TRUE;
        return;
      end_if;

      pHelpModule := pHelpModule^.pNext;
    end_while;

    pHelpCfg := pHelpCfg^.pNext;
  end_while;

END_FUNCTION

FUNCTION SafetyManager::IsCPUModule
  VAR_INPUT
    ModuleType : t_e_ModuleType;
  END_VAR
  VAR_OUTPUT
    retcode : BOOL;
  END_VAR

  case ModuleType of
    _CSCP01x,
    _SCP010,
    _SCP011,
    _SCP111,
    _SCP211,
    _SDD1300,
    _SDD1400,
    _SDD1500,
    _SDD1600:
      retcode := TRUE;
  else
    retcode := FALSE;
  end_case;

END_FUNCTION

FUNCTION SafetyManager::IsFSoEModule
  VAR_INPUT
    ModuleType 	: t_e_ModuleType;
  END_VAR
  VAR_OUTPUT
    retcode 	: BOOL;
  END_VAR

  case ModuleType of
    _SCP111,
    _SCP211,
    _SDD1300,
    _SDD1400,
    _SDD1500,
    _SDD1600,
    _ModuleWithoutConfig:
      retcode := TRUE;
  else
    retcode := FALSE;
  end_case;

END_FUNCTION

FUNCTION SafetyManager::CreateFSoEPDOs
  VAR
    pHelpConfigManager      : ^t_CfgListElem;
    pHelpConnectionManager  : ^t_FSoEConnectionDetails;
    pHelpConfigSlave        : ^t_CfgListElem;
    pHelpConnectionSlave    : ^t_FSoEConnectionDetails;
    SlavesFoundNo           : INT;
    pLastFoundSlave         : ^t_FSoEConnectionDetails;
    pLastFoundSlaveCfg      : ^t_CfgListElem;
    SortConnectionList      : BOOL;
    ConnectionsAvailable    : UINT;
    pConnectionPointerList  : pVoid;
    ActIndex                : UINT;
    pActConnection          : ^t_UdpConnection;
    i                       : UDINT;
    MandatoryUdpConMissing  : BOOL;
  END_VAR

//*****************************************************************************
//** SEARCH FOR MASTER / SLAVE PAIRS VIA SLAVE ADDRESS                       **
//*****************************************************************************

  MandatoryUdpConMissing  := FALSE;
  SortConnectionList      := FALSE;
  ConnectionsAvailable    := 0;

  // check all configs for manager connections (those contain the info about the slaves)
  pHelpConfigManager := pConfigs;
  while pHelpConfigManager do

    pHelpConnectionManager := pHelpConfigManager^.pFirstFSoEConnection;
    while pHelpConnectionManager do

      ConnectionsAvailable += 1;

      if pHelpConnectionManager^.Flags.FSoESlaveHasNoConfig & pHelpConnectionManager^.Flags.IsMaster then

        if pHelpConnectionManager^.InternalConnectionState = FCS_RESET then
          ShareSingleConnectionInfos(pHelpConnectionManager, pHelpConfigManager^.pFirstModuleCfg);
        end_if;

      // if we got a master connection => search for a match of the slaveaddress in the slave configurations
      elsif pHelpConnectionManager^.Flags.IsMaster then
        SlavesFoundNo := 0;

        if (pHelpConnectionManager^.SlavePathCompLen = UDP_COMP_PATH_LENGTH) & (pHelpConnectionManager^.pSlavePathComp^ = INTERFACE_IP_MODE) then
          // UDP Connection where we are consumer => check for it in the list of producers
          if sUdpVars.ProducerConnectionNo then
            pActConnection := #sUdpVars.paConnectionsToProducers^[0];
            for i := 0 to (sUdpVars.ProducerConnectionNo-1) do
              if (pActConnection^.IFCRC = (pHelpConnectionManager^.pSlavePathComp$^HDINT + 1)^) & (pActConnection^.IP = (pHelpConnectionManager^.pSlavePathComp$^HDINT + 5)^) then
                // check if it has to be there but isn't
                if (pActConnection^.InfoBits.IsOptional = FALSE) & (pActConnection^.InfoBits.OptionalValid = TRUE) & (pActConnection^.InfoBits.PdosInitialized = FALSE) then
                  // remember that there is something missing
                  MandatoryUdpConMissing := TRUE;
                end_if;
                exit;
              end_if;

              pActConnection += sizeof(t_UdpConnection);
            end_for;
          end_if;
        else
          pHelpConfigSlave := pConfigs;
          while pHelpConfigSlave do

            pHelpConnectionSlave := pHelpConfigSlave^.pFirstFSoEConnection;
            while pHelpConnectionSlave do
              if pHelpConnectionSlave^.Flags.IsMaster = FALSE then
                if (pHelpConnectionManager^.SlaveAddress) &
                   (pHelpConnectionManager^.SlaveAddress = pHelpConnectionSlave^.SlaveAddress) then
                  // check if it's an internal interface frame
                  if pHelpConnectionManager^.Flags.IsInterfaceConnection & pHelpConnectionSlave^.Flags.IsInterfaceConnection then
                    // check if the connection is still available
                    if pHelpConnectionSlave^.InternalConnectionState = FCS_RESET then
                      pLastFoundSlave     := pHelpConnectionSlave;
                      pLastFoundSlaveCfg  := pHelpConfigSlave;

                      // mark as internal interface frame
                      SlavesFoundNo := -1;

                      // exit both loops
                      pHelpConfigSlave := NIL;
                      exit;
                    end_if;
                  else
                    SlavesFoundNo       += 1;
                    pLastFoundSlave     := pHelpConnectionSlave;
                    pLastFoundSlaveCfg  := pHelpConfigSlave;
                  end_if;
                end_if;
              end_if;

              pHelpConnectionSlave := pHelpConnectionSlave^.pNext;
            end_while;

            if pHelpConfigSlave then
              pHelpConfigSlave := pHelpConfigSlave^.pNext;
            end_if;
          end_while;

          if SlavesFoundNo = 1 then
            // perfect, since the slave address is meant to be unique
            ShareConnectionInfos(pHelpConnectionManager, pHelpConfigManager, pLastFoundSlave, pLastFoundSlaveCfg);

          elsif SlavesFoundNo = 0 then
            // we have to search for the address in other systems which could be connected via interfaceframe
            if pFirstManagingInterfaceComponent = NIL then
              if (pHelpConnectionManager^.SlaveAddress <> 0) & (pHelpConnectionManager^.bsLogError.SlaveForMasterNotFound = FALSE) then
                LogValue("@0489 (SafetyManager::CreateFSoEPDOs) Could not find Slave for Master connection with SlaveAddress 0x{0}", Value:=pHelpConnectionManager^.SlaveAddress);
                pHelpConnectionManager^.bsLogError.SlaveForMasterNotFound := TRUE; //Only log error one time
              end_if;
            else
              SortConnectionList := TRUE;
            end_if;
          elsif SlavesFoundNo = -1 then
            // internal interface frame => add it to the list for SDO routing
            AddInternalIFFSoE(pHelpConnectionManager, pHelpConfigManager, pLastFoundSlave, pLastFoundSlaveCfg);
          else
            if pHelpConnectionManager^.bsLogError.MoreThan1SlaveFound = FALSE then
              LogValue("@048A (SafetyManager::CreateFSoEPDOs) Found more than 1 Slave for Master connection with SlaveAddress 0x{0}! Slave Address must be unique!", Value:=pHelpConnectionManager^.SlaveAddress);
              pHelpConnectionManager^.bsLogError.MoreThan1SlaveFound := TRUE; //Only log error one time
            end_if;
          end_if;
        end_if;
      else
        if pHelpConnectionManager^.Flags.IsInterfaceConnection then
          if pFirstManagingInterfaceComponent then
            SortConnectionList := TRUE;
          end_if;

          // check if we can get an interface crc from the config
          if pHelpConfigManager^.pFirstModuleCfg & (pHelpConfigManager^.pFirstModuleCfg^.ModuleInfo.SafetyNbr = pHelpConnectionManager^.OwnerSafetyNbr) then
            // store the interface CRC (to send it to the other domain later)
            if pHelpConnectionManager^.pSlavePathComp = NIL then
              pHelpConnectionManager^.pSlavePathComp$pVoid := To_StdLib.Malloc(size:=8);

              if pHelpConnectionManager^.pSlavePathComp then
                // generate a compressed path (IF CRC)
                _memset(dest:=pHelpConnectionManager^.pSlavePathComp, usByte:=16#FF, cntr:=8);
                pHelpConnectionManager^.pSlavePathComp^$USINT := 3;
                _memcpy(ptr1:=pHelpConnectionManager^.pSlavePathComp + 1, ptr2:=#pHelpConfigManager^.pFirstModuleCfg^.ModuleInfo.InterfaceCRC, cntr:=sizeof(HDINT));
                pHelpConnectionManager^.SlavePathCompLen := 8;
              else
                LogError("@048B (SafetyManager::CreateFSoEPDOs) Failed to allocate memory for an interface CRC!");
              end_if;
            end_if;
          end_if;
        end_if;
      end_if;

      pHelpConnectionManager := pHelpConnectionManager^.pNext;
    end_while;

    pHelpConfigManager := pHelpConfigManager^.pNext;
  end_while;

  if MandatoryUdpConMissing then
    // don't set b_AllLocalSlaveAddressesValid to TRUE, we need to keep waiting
    return;
  end_if;

  // check if we got all slave addresses of local configs
  CheckLocalSlaveAddresses();

  // reset pointer
  pSortedConnections := NIL;

  // there are interface connections => sort the list by slave address to ensure correct order in memory
  if SortConnectionList | (ConnectionsAvailable & (b_AllLocalSlaveAddressesValid = FALSE)) then
    // first we need a pointer list of connection (not linked) with 4 byte entries
    pConnectionPointerList := To_StdLib.Malloc(size:=ConnectionsAvailable * sizeof(pVoid));

    if pConnectionPointerList = NIL then
      LogError("@048C (SafetyManager::CreateFSoEPDOs) Failed to allocate memory for sorting the FSoE connections!");
      return;
    end_if;

    // store the pointers of all connections into the array
    ActIndex := 0;
    pHelpConfigManager := pConfigs;
    while pHelpConfigManager do

      pHelpConnectionManager := pHelpConfigManager^.pFirstFSoEConnection;
      while pHelpConnectionManager do
        (pConnectionPointerList + ActIndex * sizeof(pVoid))^$^t_FSoEConnectionDetails := pHelpConnectionManager;

        ActIndex                += 1;
        pHelpConnectionManager  := pHelpConnectionManager^.pNext;
      end_while;

      pHelpConfigManager := pHelpConfigManager^.pNext;
    end_while;

    // now that we got our linear memory to sort => do it
    MySort(src:=pConnectionPointerList$^USINT, no:=ActIndex, itemsize:=sizeof(pVoid), sortfunct:=#ConnectionSort());

    // create the new sorted linked list
    pSortedConnections := pConnectionPointerList^$^t_FSoEConnectionDetails;
    pHelpConnectionManager := pSortedConnections;

    // we already have the first connection at the pSortedConnections;
    for ActIndex := 1 to ConnectionsAvailable-1 do
      pHelpConnectionManager^.pNextSorted := (pConnectionPointerList + ActIndex * sizeof(pVoid))^$^t_FSoEConnectionDetails;
      pHelpConnectionManager := pHelpConnectionManager^.pNextSorted;
    end_for;

    To_StdLib.Free(mptr:=pConnectionPointerList);
    // now we can access the connection in order of the slave address via pSortedConnections
  end_if;

END_FUNCTION

FUNCTION SafetyManager::ShareConnectionInfos
  VAR_INPUT
    pMasterConnection 	: ^t_FSoEConnectionDetails;
    pMasterConfig 	: ^t_CfgListElem;
    pSlaveConnection 	: ^t_FSoEConnectionDetails;
    pSlaveConfig 	: ^t_CfgListElem;
  END_VAR
  VAR
    pHelpSafety   : ^t_SafetyComponent;
    pMasterSafety : ^t_SafetyComponent;
    pSlaveSafety  : ^t_SafetyComponent;
    MyPara 	      : CmdStruct;
    MyResult	    : results;
    pPDOReadData  : pVoid;
    i             : UDINT;
    IsInList      : BOOL;
  END_VAR

//*****************************************************************************
//** TELL THE MODULES WHAT DATA TO COPY IN REALTIME                          **
//*****************************************************************************

  pMasterSafety := NIL;
  pSlaveSafety  := NIL;

  pHelpSafety := pFirstSafetyComponent;
  while pHelpSafety do

    if pHelpSafety^.SafetyNbr & (pHelpSafety^.SafetyNbr = pMasterConfig^.SafetyNbr) then
      pMasterSafety := pHelpSafety;
      exit;
    end_if;

    pHelpSafety := pHelpSafety^.pNext;
  end_while;

  pHelpSafety := pFirstSafetyComponent;
  while pHelpSafety do

    if pHelpSafety^.SafetyNbr & (pHelpSafety^.SafetyNbr = pSlaveConfig^.SafetyNbr) then
      pSlaveSafety := pHelpSafety;
      exit;
    end_if;

    pHelpSafety := pHelpSafety^.pNext;
  end_while;

  // if we found the safety modules who are keeping the configs => tell them what to copy
  if pMasterSafety & pSlaveSafety then
    // check for matching hardware paths
    if (pMasterConnection^.pSlavePath^ <> pSlaveSafety^.pPath^) |
       (To_StdLib.MemCmp(pSlaveSafety^.pPath + 1, pMasterConnection^.pSlavePath + 2, pSlaveSafety^.pPath^) <> 0) then
      LogError("@048D (SafetyManager::ShareConnectionInfos) Error! The hardware path of the master connection doesn't match the hw path");
      LogValue(" of the slave module with the corresponding slave address (Slave Address 0x{0} and ConnectionID 0x{1})!", Value:=pMasterConnection^.SlaveAddress, Value2:=pMasterConnection^.ConnectionID);
      return;
    end_if;

    // check for equal sizes
    if (pMasterConnection^.MasterReadSize <> pSlaveConnection^.MasterReadSize) |
       (pMasterConnection^.MasterWriteSize <> pSlaveConnection^.MasterWriteSize) then
      LogError("@048E (SafetyManager::ShareConnectionInfos) Error! The sizes of master and slave connection");
      LogValue(" do not match for Slave Address 0x{0} and ConnectionID 0x{1}!", Value:=pMasterConnection^.SlaveAddress, Value2:=pMasterConnection^.ConnectionID);
      return;
    end_if;

    // we start with the safe outputs: get the data pointer from the master and give it to the slave
    MyPara.uiCmd    := CMD_SM_ADD_OUTPUT_PDO;
    MyResult.uiLng  := 0;
    pMasterSafety^.pThis^.NewInst(#MyPara, #MyResult);

    if MyResult.uiLng <> 4 then
      LogError("@048F (SafetyManager::ShareConnectionInfos) Invalid return value when asking the master safety module for it's pointer to the PDO read data!");
      return;
    end_if;

    pPDOReadData := MyResult.aData[0]$pVoid;

#ifdef SAFETY_DEBUG_LOGGING_ACTIVATED
#pragma message("RamAnd 20.11.2014 16:41 \ testweise mapping loggen")
    LogValue("@DBG (SafetyManager::ShareConnectionInfos) ConnectionID: {0}, SlaveAddress: {1}", Value:=pMasterConnection^.ConnectionID, Value2:=pMasterConnection^.SlaveAddress);
    LogValue("@DBG (SafetyManager::ShareConnectionInfos) MasterSafetyNbr: {0}, SlaveSafetyNbr: {1}", Value:=pMasterConnection^.OwnerSafetyNbr, Value2:=pSlaveConnection^.OwnerSafetyNbr);
    LogValue("@DBG (SafetyManager::ShareConnectionInfos) MasterReadOffset: {0}, MasterReadSize: {1}, SlaveWriteOffset: {2}", Value:=pMasterConnection^.MasterReadOffset, Value2:=pMasterConnection^.MasterReadSize, Value3 := pSlaveConnection^.SlaveWriteOffset);
#endif

    // check if it's in the list
    IsInList := FALSE;
    if FSoEInputPDONo then
      for i := 0 to (FSoEInputPDONo-1) do
        // check if the memory is already in the list for this slave safety module
        if ((aFSoEInputPDOs[i].pSafety = pSlaveSafety) & (aFSoEInputPDOs[i].pMem = pPDOReadData$DINT + pMasterConnection^.MasterReadOffset)) then
          // if we found it => skip adding the PDO to the module
          IsInList := TRUE;
        end_if;
      end_for;
    end_if;

    if IsInList = FALSE then
      MyPara.uiCmd    := CMD_SM_ADD_INPUT_PDO;
      MyPara.aPara[0] := pPDOReadData$DINT + pMasterConnection^.MasterReadOffset;
      MyPara.aPara[2] := pMasterConnection^.OwnerSafetyNbr$DINT;
      MyPara.aPara[3] := pMasterConnection^.MasterReadSize;
      MyPara.aPara[4] := pMasterSafety^.InfoBits.IsOptional;
      MyPara.aPara[7] := pSlaveConnection^.SlaveWriteOffset;
      MyPara.aPara[8] := SM_IF_VALIDITY_MARK$DINT;
      MyPara.aPara[9] := pMasterConnection^.Flags.IsInterfaceConnection;
      pSlaveSafety^.pThis^.NewInst(#MyPara, #MyResult);

      if FSoEInputPDONo < MAX_FSOE_CONNECTIONS then
        aFSoEInputPDOs[FSoEInputPDONo].pSafety    := pSlaveSafety;
        aFSoEInputPDOs[FSoEInputPDONo].pMem       := MyPara.aPara[0];
        FSoEInputPDONo += 1;
      else
        LogValue("@0490 (SafetyManager::ShareConnectionInfos) Maximum limit of allowed FSoE input Frames exceeded (0x{0})", Value:=MAX_FSOE_CONNECTIONS);
      end_if;
    end_if;

    // safe inputs: get the data pointer from the slave and give it to the master
    MyPara.uiCmd    := CMD_SM_ADD_OUTPUT_PDO;
    MyResult.uiLng  := 0;
    pSlaveSafety^.pThis^.NewInst(#MyPara, #MyResult);

    if MyResult.uiLng <> 4 then
      LogError("@0491 (SafetyManager::ShareConnectionInfos) Invalid return value when asking the slave safety module for it's pointer to the PDO read data!");
      return;
    end_if;

    pPDOReadData := MyResult.aData[0]$pVoid;

#ifdef SAFETY_DEBUG_LOGGING_ACTIVATED
#pragma message("RamAnd 20.11.2014 16:41 \ testweise mapping loggen")
    LogValue("@DBG (SafetyManager::ShareConnectionInfos) SlaveReadOffset: {0}, SlaveReadSize: {1}, MasterWriteOffset: {2}", Value:=pSlaveConnection^.SlaveReadOffset, Value2:=pMasterConnection^.MasterWriteSize, Value3 := pMasterConnection^.MasterWriteOffset);
#endif

    // check if it's in the list
    IsInList := FALSE;
    if FSoEInputPDONo then
      for i := 0 to (FSoEInputPDONo-1) do
        // check if the memory is already in the list for this slave safety module
        if ((aFSoEInputPDOs[i].pSafety = pMasterSafety)  & (aFSoEInputPDOs[i].pMem = pPDOReadData$DINT + pSlaveConnection^.SlaveReadOffset)) then
          // if we found it => skip adding the PDO to the module
          IsInList := TRUE;
        end_if;
      end_for;
    end_if;

    if IsInList = FALSE then

      MyPara.uiCmd    := CMD_SM_ADD_INPUT_PDO;
      MyPara.aPara[0] := pPDOReadData$DINT + pSlaveConnection^.SlaveReadOffset;
      MyPara.aPara[2] := pSlaveConnection^.OwnerSafetyNbr$DINT;
      MyPara.aPara[3] := pMasterConnection^.MasterWriteSize;
      MyPara.aPara[4] := pSlaveSafety^.InfoBits.IsOptional;
      MyPara.aPara[7] := pMasterConnection^.MasterWriteOffset;
      MyPara.aPara[8] := 0;
      MyPara.aPara[9] := 0;
      pMasterSafety^.pThis^.NewInst(#MyPara, #MyResult);

      if FSoEInputPDONo < MAX_FSOE_CONNECTIONS then
        aFSoEInputPDOs[FSoEInputPDONo].pSafety    := pMasterSafety;
        aFSoEInputPDOs[FSoEInputPDONo].pMem       := MyPara.aPara[0];
        FSoEInputPDONo += 1;
      else
        LogValue("@0490 (SafetyManager::ShareConnectionInfos) Maximum limit of allowed FSoE input Frames exceeded (0x{0})", Value:=MAX_FSOE_CONNECTIONS);
      end_if;
    end_if;
  end_if;

END_FUNCTION

FUNCTION MyXSort VAR_INPUT p1:^void; p2:^void; END_VAR VAR_OUTPUT retcode : dint; END_VAR;

FUNCTION SafetyManager::MySort
  VAR_INPUT
    src 	: ^USINT;
    no 	: UDINT;
    itemsize 	: UDINT;
    sortfunct 	: ^void;
  END_VAR
  VAR_OUTPUT
    retcode 	: BOOL;
  END_VAR
  var
    tmp, hp : ^DINT;
    mx, nx, wx, parent, child, max, i : dint;
    spuf : array[0..127] of dint;
  end_var

  retcode := false;

  // work faster with the pointer list (no memcopy used)
  if itemsize = 4 then
    nx      := to_dint(no);
    mx      := (nx + 6) / 8;
    src     := src;
    tmp     := #spuf[0];
    retcode := true;

    while(1) do
      if(mx) then
        mx     -= 1;
        parent := mx;
        tmp^ := (src$^DINT + (parent$udint*4))^;
      else
        nx -= 1;
        if(nx) then
          hp := src + (nx$udint*4);
          tmp^ := hp^;
          hp^ := (src$^DINT)^;
          parent := 0;
        else
          exit;
        end_if;
      end_if;
